(* IEC 61131-3 sources: sis-interlock-demo/tests/POUs/Generated/FB_VoteTruth_Test, 83 files *)

(* ---- FB_VoteTruth_Test.decl.st ---- *)
// AUTO-GENERATED by cemgen 1.0.0 — не редактировать: правьте матрицу и запустите
//   python -m cemgen generate <файл матрицы .csv или .xlsx>
// Матрица: SIS-V101-CEM, объект V-101, ревизия B от 2026-10-19, SHA-256 сетки df2ed4841a9453ca
// Назначение: набор coUnit: таблицы истинности голосования — F_VoteEval и FB_Voting по всем схемам,
//             политикам деградации и видам входа (DESIGN.md, 12.2). Экземпляр — GVL_TestsGenerated.
// Автор:      kr0nsch; код — генератор cemgen
// Версия:     1.0.0
// Документ:   docs/DESIGN.md, раздел «10. Генератор cemgen»; docs/cause_effect_matrix.md
// ВНИМАНИЕ:   код демонстрационный и не предназначен для систем безопасности. Реальная ПАЗ требует
//             определения SIL, сертифицированных аппаратных и программных средств и валидации по
//             ГОСТ Р МЭК 61511.
FUNCTION_BLOCK FB_VoteTruth_Test EXTENDS coUnit.FB_TestSuite
VAR
END_VAR

(* ---- ArchIndex.method.decl.st ---- *)
// AUTO-GENERATED by cemgen 1.0.0 — не редактировать: правьте матрицу и запустите
//   python -m cemgen generate <файл матрицы .csv или .xlsx>
// Матрица: SIS-V101-CEM, объект V-101, ревизия B от 2026-10-19, SHA-256 сетки df2ed4841a9453ca
// Назначение: вспомогательный метод набора FB_VoteTruth_Test.
// Автор:      kr0nsch; код — генератор cemgen
// Версия:     1.0.0
// Документ:   docs/DESIGN.md, раздел «10. Генератор cemgen»; docs/cause_effect_matrix.md
// ВНИМАНИЕ:   код демонстрационный и не предназначен для систем безопасности. Реальная ПАЗ требует
//             определения SIL, сертифицированных аппаратных и программных средств и валидации по
//             ГОСТ Р МЭК 61511.
// Индекс схемы в байте таблицы: 0 None, 1 1oo1, 2 1oo2, 3 2oo2, 4 2oo3, 5 ForcedTrip.
METHOD PRIVATE ArchIndex : BYTE
VAR_INPUT
    eArch : E_VoteArch;   // действующая схема
END_VAR

(* ---- ArchIndex.method.impl.st ---- *)
// AUTO-GENERATED by cemgen 1.0.0 — не редактировать: правьте матрицу и запустите
//   python -m cemgen generate <файл матрицы .csv или .xlsx>
// Матрица: SIS-V101-CEM, объект V-101, ревизия B от 2026-10-19, SHA-256 сетки df2ed4841a9453ca
CASE eArch OF
    E_VoteArch.Vote1oo1:
        ArchIndex := 1;
    E_VoteArch.Vote1oo2:
        ArchIndex := 2;
    E_VoteArch.Vote2oo2:
        ArchIndex := 3;
    E_VoteArch.Vote2oo3:
        ArchIndex := 4;
    E_VoteArch.ForcedTrip:
        ArchIndex := 5;
ELSE
    ArchIndex := 0;
END_CASE

(* ---- EncodeEval.method.decl.st ---- *)
// AUTO-GENERATED by cemgen 1.0.0 — не редактировать: правьте матрицу и запустите
//   python -m cemgen generate <файл матрицы .csv или .xlsx>
// Матрица: SIS-V101-CEM, объект V-101, ревизия B от 2026-10-19, SHA-256 сетки df2ed4841a9453ca
// Назначение: вспомогательный метод набора FB_VoteTruth_Test.
// Автор:      kr0nsch; код — генератор cemgen
// Версия:     1.0.0
// Документ:   docs/DESIGN.md, раздел «10. Генератор cemgen»; docs/cause_effect_matrix.md
// ВНИМАНИЕ:   код демонстрационный и не предназначен для систем безопасности. Реальная ПАЗ требует
//             определения SIL, сертифицированных аппаратных и программных средств и валидации по
//             ГОСТ Р МЭК 61511.
// Байт результата F_VoteEval: бит 0 — xTrip, бит 1 — xDegraded, биты 2–4 — индекс eArchEff.
METHOD PRIVATE EncodeEval : BYTE
VAR_INPUT
    stRes : ST_VoteResult;   // результат F_VoteEval
END_VAR

(* ---- EncodeFb.method.decl.st ---- *)
// AUTO-GENERATED by cemgen 1.0.0 — не редактировать: правьте матрицу и запустите
//   python -m cemgen generate <файл матрицы .csv или .xlsx>
// Матрица: SIS-V101-CEM, объект V-101, ревизия B от 2026-10-19, SHA-256 сетки df2ed4841a9453ca
// Назначение: вспомогательный метод набора FB_VoteTruth_Test.
// Автор:      kr0nsch; код — генератор cemgen
// Версия:     1.0.0
// Документ:   docs/DESIGN.md, раздел «10. Генератор cemgen»; docs/cause_effect_matrix.md
// ВНИМАНИЕ:   код демонстрационный и не предназначен для систем безопасности. Реальная ПАЗ требует
//             определения SIL, сертифицированных аппаратных и программных средств и валидации по
//             ГОСТ Р МЭК 61511.
// Байт результата FB_Voting: как у EncodeEval, плюс биты 5–7 — байпас каналов 1–3 в состоянии Active.
METHOD PRIVATE EncodeFb : BYTE
VAR_INPUT
    xTrip : BOOL;           // выход xTrip
    stSts : ST_VotingSts;   // состояние группы
END_VAR
VAR
    uiCh : UINT;            // канал
END_VAR

(* ---- EncodeFb.method.impl.st ---- *)
// AUTO-GENERATED by cemgen 1.0.0 — не редактировать: правьте матрицу и запустите
//   python -m cemgen generate <файл матрицы .csv или .xlsx>
// Матрица: SIS-V101-CEM, объект V-101, ревизия B от 2026-10-19, SHA-256 сетки df2ed4841a9453ca
EncodeFb := BOOL_TO_BYTE(xTrip) OR SHL(BOOL_TO_BYTE(stSts.xDegraded), 1)
    OR SHL(ArchIndex(eArch := stSts.eArchEff), 2);
FOR uiCh := 1 TO GVL_Const.SIS_VOTE_CH_MAX DO
    EncodeFb := EncodeFb OR SHL(BOOL_TO_BYTE(stSts.aeBypass[uiCh] = E_BypassState.Active), 4 + uiCh);
END_FOR

(* ---- Eval1oo1DAMatchesTable.method.decl.st ---- *)
// AUTO-GENERATED by cemgen 1.0.0 — не редактировать: правьте матрицу и запустите
//   python -m cemgen generate <файл матрицы .csv или .xlsx>
// Матрица: SIS-V101-CEM, объект V-101, ревизия B от 2026-10-19, SHA-256 сетки df2ed4841a9453ca
// Назначение: тест VoteTruth_Eval1oo1DA_MatchesTable набора FB_VoteTruth_Test.
// Автор:      kr0nsch; код — генератор cemgen
// Версия:     1.0.0
// Документ:   docs/DESIGN.md, раздел «10. Генератор cemgen»; docs/cause_effect_matrix.md
// ВНИМАНИЕ:   код демонстрационный и не предназначен для систем безопасности. Реальная ПАЗ требует
//             определения SIL, сертифицированных аппаратных и программных средств и валидации по
//             ГОСТ Р МЭК 61511.
// F_VoteEval, схема 1oo1, политика DegradeAvailable: все 4 сочетаний состояний каналов (Normal,
// Demand, Invalid, Bypassed) совпадают с таблицей TT_EVAL_1OO1_DA.
METHOD PRIVATE Eval1oo1DAMatchesTable
VAR
    uiRow      : UINT;                                                    // строка таблицы
    aeCh       : ARRAY[1..GVL_Const.SIS_VOTE_CH_MAX] OF E_ChannelState;   // состояния каналов строки
    stRes      : ST_VoteResult;                                           // результат F_VoteEval
    bAct       : BYTE;                                                    // фактический байт результата
    bExp       : BYTE;                                                    // ожидаемый байт из таблицы
    xMiss      : BOOL;                                                    // строка не совпала
    xFirst     : BOOL;                                                    // первая несовпавшая строка
    uiMismatch : UINT;                                                    // несовпавших строк
    uiFirstRow : UINT;                                                    // первая несовпавшая строка
    bFirstExp  : BYTE;                                                    // ожидаемый байт первой несовпавшей строки
    bFirstAct  : BYTE;                                                    // фактический байт первой несовпавшей строки
END_VAR

(* ---- Eval1oo1DAMatchesTable.method.impl.st ---- *)
// AUTO-GENERATED by cemgen 1.0.0 — не редактировать: правьте матрицу и запустите
//   python -m cemgen generate <файл матрицы .csv или .xlsx>
// Матрица: SIS-V101-CEM, объект V-101, ревизия B от 2026-10-19, SHA-256 сетки df2ed4841a9453ca
coUnit.TEST('VoteTruth_Eval1oo1DA_MatchesTable');
FOR uiRow := 0 TO 3 DO
    RowStates(uiRow := uiRow, uiChannels := 1, aeCh := aeCh);
    stRes := F_VoteEval(eArch := E_VoteArch.Vote1oo1, ePolicy := E_DegradePolicy.DegradeAvailable,
        aeCh := aeCh);
    bAct := EncodeEval(stRes := stRes);
    bExp := GVL_VoteTruthTable.TT_EVAL_1OO1_DA[uiRow];
    xMiss := bAct <> bExp;
    xFirst := xMiss AND uiMismatch = 0;
    uiFirstRow := SEL(xFirst, uiFirstRow, uiRow);
    bFirstExp := SEL(xFirst, bFirstExp, bExp);
    bFirstAct := SEL(xFirst, bFirstAct, bAct);
    uiMismatch := uiMismatch + BOOL_TO_UINT(xMiss);
END_FOR
AssertEquals_UINT(Expected := 0, Actual := uiMismatch,
    Message := MismatchText(sTable := 'TT_EVAL_1OO1_DA', uiRow := uiFirstRow, bExpected := bFirstExp,
        bActual := bFirstAct));
coUnit.TEST_FINISHED();

(* ---- Eval1oo1DSMatchesTable.method.decl.st ---- *)
// AUTO-GENERATED by cemgen 1.0.0 — не редактировать: правьте матрицу и запустите
//   python -m cemgen generate <файл матрицы .csv или .xlsx>
// Матрица: SIS-V101-CEM, объект V-101, ревизия B от 2026-10-19, SHA-256 сетки df2ed4841a9453ca
// Назначение: тест VoteTruth_Eval1oo1DS_MatchesTable набора FB_VoteTruth_Test.
// Автор:      kr0nsch; код — генератор cemgen
// Версия:     1.0.0
// Документ:   docs/DESIGN.md, раздел «10. Генератор cemgen»; docs/cause_effect_matrix.md
// ВНИМАНИЕ:   код демонстрационный и не предназначен для систем безопасности. Реальная ПАЗ требует
//             определения SIL, сертифицированных аппаратных и программных средств и валидации по
//             ГОСТ Р МЭК 61511.
// F_VoteEval, схема 1oo1, политика DegradeSafe: все 4 сочетаний состояний каналов (Normal, Demand,
// Invalid, Bypassed) совпадают с таблицей TT_EVAL_1OO1_DS.
METHOD PRIVATE Eval1oo1DSMatchesTable
VAR
    uiRow      : UINT;                                                    // строка таблицы
    aeCh       : ARRAY[1..GVL_Const.SIS_VOTE_CH_MAX] OF E_ChannelState;   // состояния каналов строки
    stRes      : ST_VoteResult;                                           // результат F_VoteEval
    bAct       : BYTE;                                                    // фактический байт результата
    bExp       : BYTE;                                                    // ожидаемый байт из таблицы
    xMiss      : BOOL;                                                    // строка не совпала
    xFirst     : BOOL;                                                    // первая несовпавшая строка
    uiMismatch : UINT;                                                    // несовпавших строк
    uiFirstRow : UINT;                                                    // первая несовпавшая строка
    bFirstExp  : BYTE;                                                    // ожидаемый байт первой несовпавшей строки
    bFirstAct  : BYTE;                                                    // фактический байт первой несовпавшей строки
END_VAR

(* ---- Eval1oo1DSMatchesTable.method.impl.st ---- *)
// AUTO-GENERATED by cemgen 1.0.0 — не редактировать: правьте матрицу и запустите
//   python -m cemgen generate <файл матрицы .csv или .xlsx>
// Матрица: SIS-V101-CEM, объект V-101, ревизия B от 2026-10-19, SHA-256 сетки df2ed4841a9453ca
coUnit.TEST('VoteTruth_Eval1oo1DS_MatchesTable');
FOR uiRow := 0 TO 3 DO
    RowStates(uiRow := uiRow, uiChannels := 1, aeCh := aeCh);
    stRes := F_VoteEval(eArch := E_VoteArch.Vote1oo1, ePolicy := E_DegradePolicy.DegradeSafe,
        aeCh := aeCh);
    bAct := EncodeEval(stRes := stRes);
    bExp := GVL_VoteTruthTable.TT_EVAL_1OO1_DS[uiRow];
    xMiss := bAct <> bExp;
    xFirst := xMiss AND uiMismatch = 0;
    uiFirstRow := SEL(xFirst, uiFirstRow, uiRow);
    bFirstExp := SEL(xFirst, bFirstExp, bExp);
    bFirstAct := SEL(xFirst, bFirstAct, bAct);
    uiMismatch := uiMismatch + BOOL_TO_UINT(xMiss);
END_FOR
AssertEquals_UINT(Expected := 0, Actual := uiMismatch,
    Message := MismatchText(sTable := 'TT_EVAL_1OO1_DS', uiRow := uiFirstRow, bExpected := bFirstExp,
        bActual := bFirstAct));
coUnit.TEST_FINISHED();

(* ---- Eval1oo1VTMatchesTable.method.decl.st ---- *)
// AUTO-GENERATED by cemgen 1.0.0 — не редактировать: правьте матрицу и запустите
//   python -m cemgen generate <файл матрицы .csv или .xlsx>
// Матрица: SIS-V101-CEM, объект V-101, ревизия B от 2026-10-19, SHA-256 сетки df2ed4841a9453ca
// Назначение: тест VoteTruth_Eval1oo1VT_MatchesTable набора FB_VoteTruth_Test.
// Автор:      kr0nsch; код — генератор cemgen
// Версия:     1.0.0
// Документ:   docs/DESIGN.md, раздел «10. Генератор cemgen»; docs/cause_effect_matrix.md
// ВНИМАНИЕ:   код демонстрационный и не предназначен для систем безопасности. Реальная ПАЗ требует
//             определения SIL, сертифицированных аппаратных и программных средств и валидации по
//             ГОСТ Р МЭК 61511.
// F_VoteEval, схема 1oo1, политика VoteTrip: все 4 сочетаний состояний каналов (Normal, Demand,
// Invalid, Bypassed) совпадают с таблицей TT_EVAL_1OO1_VT.
METHOD PRIVATE Eval1oo1VTMatchesTable
VAR
    uiRow      : UINT;                                                    // строка таблицы
    aeCh       : ARRAY[1..GVL_Const.SIS_VOTE_CH_MAX] OF E_ChannelState;   // состояния каналов строки
    stRes      : ST_VoteResult;                                           // результат F_VoteEval
    bAct       : BYTE;                                                    // фактический байт результата
    bExp       : BYTE;                                                    // ожидаемый байт из таблицы
    xMiss      : BOOL;                                                    // строка не совпала
    xFirst     : BOOL;                                                    // первая несовпавшая строка
    uiMismatch : UINT;                                                    // несовпавших строк
    uiFirstRow : UINT;                                                    // первая несовпавшая строка
    bFirstExp  : BYTE;                                                    // ожидаемый байт первой несовпавшей строки
    bFirstAct  : BYTE;                                                    // фактический байт первой несовпавшей строки
END_VAR

(* ---- Eval1oo1VTMatchesTable.method.impl.st ---- *)
// AUTO-GENERATED by cemgen 1.0.0 — не редактировать: правьте матрицу и запустите
//   python -m cemgen generate <файл матрицы .csv или .xlsx>
// Матрица: SIS-V101-CEM, объект V-101, ревизия B от 2026-10-19, SHA-256 сетки df2ed4841a9453ca
coUnit.TEST('VoteTruth_Eval1oo1VT_MatchesTable');
FOR uiRow := 0 TO 3 DO
    RowStates(uiRow := uiRow, uiChannels := 1, aeCh := aeCh);
    stRes := F_VoteEval(eArch := E_VoteArch.Vote1oo1, ePolicy := E_DegradePolicy.VoteTrip,
        aeCh := aeCh);
    bAct := EncodeEval(stRes := stRes);
    bExp := GVL_VoteTruthTable.TT_EVAL_1OO1_VT[uiRow];
    xMiss := bAct <> bExp;
    xFirst := xMiss AND uiMismatch = 0;
    uiFirstRow := SEL(xFirst, uiFirstRow, uiRow);
    bFirstExp := SEL(xFirst, bFirstExp, bExp);
    bFirstAct := SEL(xFirst, bFirstAct, bAct);
    uiMismatch := uiMismatch + BOOL_TO_UINT(xMiss);
END_FOR
AssertEquals_UINT(Expected := 0, Actual := uiMismatch,
    Message := MismatchText(sTable := 'TT_EVAL_1OO1_VT', uiRow := uiFirstRow, bExpected := bFirstExp,
        bActual := bFirstAct));
coUnit.TEST_FINISHED();

(* ---- Eval1oo2DAMatchesTable.method.decl.st ---- *)
// AUTO-GENERATED by cemgen 1.0.0 — не редактировать: правьте матрицу и запустите
//   python -m cemgen generate <файл матрицы .csv или .xlsx>
// Матрица: SIS-V101-CEM, объект V-101, ревизия B от 2026-10-19, SHA-256 сетки df2ed4841a9453ca
// Назначение: тест VoteTruth_Eval1oo2DA_MatchesTable набора FB_VoteTruth_Test.
// Автор:      kr0nsch; код — генератор cemgen
// Версия:     1.0.0
// Документ:   docs/DESIGN.md, раздел «10. Генератор cemgen»; docs/cause_effect_matrix.md
// ВНИМАНИЕ:   код демонстрационный и не предназначен для систем безопасности. Реальная ПАЗ требует
//             определения SIL, сертифицированных аппаратных и программных средств и валидации по
//             ГОСТ Р МЭК 61511.
// F_VoteEval, схема 1oo2, политика DegradeAvailable: все 16 сочетаний состояний каналов (Normal,
// Demand, Invalid, Bypassed) совпадают с таблицей TT_EVAL_1OO2_DA.
METHOD PRIVATE Eval1oo2DAMatchesTable
VAR
    uiRow      : UINT;                                                    // строка таблицы
    aeCh       : ARRAY[1..GVL_Const.SIS_VOTE_CH_MAX] OF E_ChannelState;   // состояния каналов строки
    stRes      : ST_VoteResult;                                           // результат F_VoteEval
    bAct       : BYTE;                                                    // фактический байт результата
    bExp       : BYTE;                                                    // ожидаемый байт из таблицы
    xMiss      : BOOL;                                                    // строка не совпала
    xFirst     : BOOL;                                                    // первая несовпавшая строка
    uiMismatch : UINT;                                                    // несовпавших строк
    uiFirstRow : UINT;                                                    // первая несовпавшая строка
    bFirstExp  : BYTE;                                                    // ожидаемый байт первой несовпавшей строки
    bFirstAct  : BYTE;                                                    // фактический байт первой несовпавшей строки
END_VAR

(* ---- Eval1oo2DAMatchesTable.method.impl.st ---- *)
// AUTO-GENERATED by cemgen 1.0.0 — не редактировать: правьте матрицу и запустите
//   python -m cemgen generate <файл матрицы .csv или .xlsx>
// Матрица: SIS-V101-CEM, объект V-101, ревизия B от 2026-10-19, SHA-256 сетки df2ed4841a9453ca
coUnit.TEST('VoteTruth_Eval1oo2DA_MatchesTable');
FOR uiRow := 0 TO 15 DO
    RowStates(uiRow := uiRow, uiChannels := 2, aeCh := aeCh);
    stRes := F_VoteEval(eArch := E_VoteArch.Vote1oo2, ePolicy := E_DegradePolicy.DegradeAvailable,
        aeCh := aeCh);
    bAct := EncodeEval(stRes := stRes);
    bExp := GVL_VoteTruthTable.TT_EVAL_1OO2_DA[uiRow];
    xMiss := bAct <> bExp;
    xFirst := xMiss AND uiMismatch = 0;
    uiFirstRow := SEL(xFirst, uiFirstRow, uiRow);
    bFirstExp := SEL(xFirst, bFirstExp, bExp);
    bFirstAct := SEL(xFirst, bFirstAct, bAct);
    uiMismatch := uiMismatch + BOOL_TO_UINT(xMiss);
END_FOR
AssertEquals_UINT(Expected := 0, Actual := uiMismatch,
    Message := MismatchText(sTable := 'TT_EVAL_1OO2_DA', uiRow := uiFirstRow, bExpected := bFirstExp,
        bActual := bFirstAct));
coUnit.TEST_FINISHED();

(* ---- Eval1oo2DSMatchesTable.method.decl.st ---- *)
// AUTO-GENERATED by cemgen 1.0.0 — не редактировать: правьте матрицу и запустите
//   python -m cemgen generate <файл матрицы .csv или .xlsx>
// Матрица: SIS-V101-CEM, объект V-101, ревизия B от 2026-10-19, SHA-256 сетки df2ed4841a9453ca
// Назначение: тест VoteTruth_Eval1oo2DS_MatchesTable набора FB_VoteTruth_Test.
// Автор:      kr0nsch; код — генератор cemgen
// Версия:     1.0.0
// Документ:   docs/DESIGN.md, раздел «10. Генератор cemgen»; docs/cause_effect_matrix.md
// ВНИМАНИЕ:   код демонстрационный и не предназначен для систем безопасности. Реальная ПАЗ требует
//             определения SIL, сертифицированных аппаратных и программных средств и валидации по
//             ГОСТ Р МЭК 61511.
// F_VoteEval, схема 1oo2, политика DegradeSafe: все 16 сочетаний состояний каналов (Normal, Demand,
// Invalid, Bypassed) совпадают с таблицей TT_EVAL_1OO2_DS.
METHOD PRIVATE Eval1oo2DSMatchesTable
VAR
    uiRow      : UINT;                                                    // строка таблицы
    aeCh       : ARRAY[1..GVL_Const.SIS_VOTE_CH_MAX] OF E_ChannelState;   // состояния каналов строки
    stRes      : ST_VoteResult;                                           // результат F_VoteEval
    bAct       : BYTE;                                                    // фактический байт результата
    bExp       : BYTE;                                                    // ожидаемый байт из таблицы
    xMiss      : BOOL;                                                    // строка не совпала
    xFirst     : BOOL;                                                    // первая несовпавшая строка
    uiMismatch : UINT;                                                    // несовпавших строк
    uiFirstRow : UINT;                                                    // первая несовпавшая строка
    bFirstExp  : BYTE;                                                    // ожидаемый байт первой несовпавшей строки
    bFirstAct  : BYTE;                                                    // фактический байт первой несовпавшей строки
END_VAR

(* ---- Eval1oo2DSMatchesTable.method.impl.st ---- *)
// AUTO-GENERATED by cemgen 1.0.0 — не редактировать: правьте матрицу и запустите
//   python -m cemgen generate <файл матрицы .csv или .xlsx>
// Матрица: SIS-V101-CEM, объект V-101, ревизия B от 2026-10-19, SHA-256 сетки df2ed4841a9453ca
coUnit.TEST('VoteTruth_Eval1oo2DS_MatchesTable');
FOR uiRow := 0 TO 15 DO
    RowStates(uiRow := uiRow, uiChannels := 2, aeCh := aeCh);
    stRes := F_VoteEval(eArch := E_VoteArch.Vote1oo2, ePolicy := E_DegradePolicy.DegradeSafe,
        aeCh := aeCh);
    bAct := EncodeEval(stRes := stRes);
    bExp := GVL_VoteTruthTable.TT_EVAL_1OO2_DS[uiRow];
    xMiss := bAct <> bExp;
    xFirst := xMiss AND uiMismatch = 0;
    uiFirstRow := SEL(xFirst, uiFirstRow, uiRow);
    bFirstExp := SEL(xFirst, bFirstExp, bExp);
    bFirstAct := SEL(xFirst, bFirstAct, bAct);
    uiMismatch := uiMismatch + BOOL_TO_UINT(xMiss);
END_FOR
AssertEquals_UINT(Expected := 0, Actual := uiMismatch,
    Message := MismatchText(sTable := 'TT_EVAL_1OO2_DS', uiRow := uiFirstRow, bExpected := bFirstExp,
        bActual := bFirstAct));
coUnit.TEST_FINISHED();

(* ---- Eval1oo2VTMatchesTable.method.decl.st ---- *)
// AUTO-GENERATED by cemgen 1.0.0 — не редактировать: правьте матрицу и запустите
//   python -m cemgen generate <файл матрицы .csv или .xlsx>
// Матрица: SIS-V101-CEM, объект V-101, ревизия B от 2026-10-19, SHA-256 сетки df2ed4841a9453ca
// Назначение: тест VoteTruth_Eval1oo2VT_MatchesTable набора FB_VoteTruth_Test.
// Автор:      kr0nsch; код — генератор cemgen
// Версия:     1.0.0
// Документ:   docs/DESIGN.md, раздел «10. Генератор cemgen»; docs/cause_effect_matrix.md
// ВНИМАНИЕ:   код демонстрационный и не предназначен для систем безопасности. Реальная ПАЗ требует
//             определения SIL, сертифицированных аппаратных и программных средств и валидации по
//             ГОСТ Р МЭК 61511.
// F_VoteEval, схема 1oo2, политика VoteTrip: все 16 сочетаний состояний каналов (Normal, Demand,
// Invalid, Bypassed) совпадают с таблицей TT_EVAL_1OO2_VT.
METHOD PRIVATE Eval1oo2VTMatchesTable
VAR
    uiRow      : UINT;                                                    // строка таблицы
    aeCh       : ARRAY[1..GVL_Const.SIS_VOTE_CH_MAX] OF E_ChannelState;   // состояния каналов строки
    stRes      : ST_VoteResult;                                           // результат F_VoteEval
    bAct       : BYTE;                                                    // фактический байт результата
    bExp       : BYTE;                                                    // ожидаемый байт из таблицы
    xMiss      : BOOL;                                                    // строка не совпала
    xFirst     : BOOL;                                                    // первая несовпавшая строка
    uiMismatch : UINT;                                                    // несовпавших строк
    uiFirstRow : UINT;                                                    // первая несовпавшая строка
    bFirstExp  : BYTE;                                                    // ожидаемый байт первой несовпавшей строки
    bFirstAct  : BYTE;                                                    // фактический байт первой несовпавшей строки
END_VAR

(* ---- Eval1oo2VTMatchesTable.method.impl.st ---- *)
// AUTO-GENERATED by cemgen 1.0.0 — не редактировать: правьте матрицу и запустите
//   python -m cemgen generate <файл матрицы .csv или .xlsx>
// Матрица: SIS-V101-CEM, объект V-101, ревизия B от 2026-10-19, SHA-256 сетки df2ed4841a9453ca
coUnit.TEST('VoteTruth_Eval1oo2VT_MatchesTable');
FOR uiRow := 0 TO 15 DO
    RowStates(uiRow := uiRow, uiChannels := 2, aeCh := aeCh);
    stRes := F_VoteEval(eArch := E_VoteArch.Vote1oo2, ePolicy := E_DegradePolicy.VoteTrip,
        aeCh := aeCh);
    bAct := EncodeEval(stRes := stRes);
    bExp := GVL_VoteTruthTable.TT_EVAL_1OO2_VT[uiRow];
    xMiss := bAct <> bExp;
    xFirst := xMiss AND uiMismatch = 0;
    uiFirstRow := SEL(xFirst, uiFirstRow, uiRow);
    bFirstExp := SEL(xFirst, bFirstExp, bExp);
    bFirstAct := SEL(xFirst, bFirstAct, bAct);
    uiMismatch := uiMismatch + BOOL_TO_UINT(xMiss);
END_FOR
AssertEquals_UINT(Expected := 0, Actual := uiMismatch,
    Message := MismatchText(sTable := 'TT_EVAL_1OO2_VT', uiRow := uiFirstRow, bExpected := bFirstExp,
        bActual := bFirstAct));
coUnit.TEST_FINISHED();

(* ---- Eval2oo2DAMatchesTable.method.decl.st ---- *)
// AUTO-GENERATED by cemgen 1.0.0 — не редактировать: правьте матрицу и запустите
//   python -m cemgen generate <файл матрицы .csv или .xlsx>
// Матрица: SIS-V101-CEM, объект V-101, ревизия B от 2026-10-19, SHA-256 сетки df2ed4841a9453ca
// Назначение: тест VoteTruth_Eval2oo2DA_MatchesTable набора FB_VoteTruth_Test.
// Автор:      kr0nsch; код — генератор cemgen
// Версия:     1.0.0
// Документ:   docs/DESIGN.md, раздел «10. Генератор cemgen»; docs/cause_effect_matrix.md
// ВНИМАНИЕ:   код демонстрационный и не предназначен для систем безопасности. Реальная ПАЗ требует
//             определения SIL, сертифицированных аппаратных и программных средств и валидации по
//             ГОСТ Р МЭК 61511.
// F_VoteEval, схема 2oo2, политика DegradeAvailable: все 16 сочетаний состояний каналов (Normal,
// Demand, Invalid, Bypassed) совпадают с таблицей TT_EVAL_2OO2_DA.
METHOD PRIVATE Eval2oo2DAMatchesTable
VAR
    uiRow      : UINT;                                                    // строка таблицы
    aeCh       : ARRAY[1..GVL_Const.SIS_VOTE_CH_MAX] OF E_ChannelState;   // состояния каналов строки
    stRes      : ST_VoteResult;                                           // результат F_VoteEval
    bAct       : BYTE;                                                    // фактический байт результата
    bExp       : BYTE;                                                    // ожидаемый байт из таблицы
    xMiss      : BOOL;                                                    // строка не совпала
    xFirst     : BOOL;                                                    // первая несовпавшая строка
    uiMismatch : UINT;                                                    // несовпавших строк
    uiFirstRow : UINT;                                                    // первая несовпавшая строка
    bFirstExp  : BYTE;                                                    // ожидаемый байт первой несовпавшей строки
    bFirstAct  : BYTE;                                                    // фактический байт первой несовпавшей строки
END_VAR

(* ---- Eval2oo2DAMatchesTable.method.impl.st ---- *)
// AUTO-GENERATED by cemgen 1.0.0 — не редактировать: правьте матрицу и запустите
//   python -m cemgen generate <файл матрицы .csv или .xlsx>
// Матрица: SIS-V101-CEM, объект V-101, ревизия B от 2026-10-19, SHA-256 сетки df2ed4841a9453ca
coUnit.TEST('VoteTruth_Eval2oo2DA_MatchesTable');
FOR uiRow := 0 TO 15 DO
    RowStates(uiRow := uiRow, uiChannels := 2, aeCh := aeCh);
    stRes := F_VoteEval(eArch := E_VoteArch.Vote2oo2, ePolicy := E_DegradePolicy.DegradeAvailable,
        aeCh := aeCh);
    bAct := EncodeEval(stRes := stRes);
    bExp := GVL_VoteTruthTable.TT_EVAL_2OO2_DA[uiRow];
    xMiss := bAct <> bExp;
    xFirst := xMiss AND uiMismatch = 0;
    uiFirstRow := SEL(xFirst, uiFirstRow, uiRow);
    bFirstExp := SEL(xFirst, bFirstExp, bExp);
    bFirstAct := SEL(xFirst, bFirstAct, bAct);
    uiMismatch := uiMismatch + BOOL_TO_UINT(xMiss);
END_FOR
AssertEquals_UINT(Expected := 0, Actual := uiMismatch,
    Message := MismatchText(sTable := 'TT_EVAL_2OO2_DA', uiRow := uiFirstRow, bExpected := bFirstExp,
        bActual := bFirstAct));
coUnit.TEST_FINISHED();

(* ---- Eval2oo2DSMatchesTable.method.decl.st ---- *)
// AUTO-GENERATED by cemgen 1.0.0 — не редактировать: правьте матрицу и запустите
//   python -m cemgen generate <файл матрицы .csv или .xlsx>
// Матрица: SIS-V101-CEM, объект V-101, ревизия B от 2026-10-19, SHA-256 сетки df2ed4841a9453ca
// Назначение: тест VoteTruth_Eval2oo2DS_MatchesTable набора FB_VoteTruth_Test.
// Автор:      kr0nsch; код — генератор cemgen
// Версия:     1.0.0
// Документ:   docs/DESIGN.md, раздел «10. Генератор cemgen»; docs/cause_effect_matrix.md
// ВНИМАНИЕ:   код демонстрационный и не предназначен для систем безопасности. Реальная ПАЗ требует
//             определения SIL, сертифицированных аппаратных и программных средств и валидации по
//             ГОСТ Р МЭК 61511.
// F_VoteEval, схема 2oo2, политика DegradeSafe: все 16 сочетаний состояний каналов (Normal, Demand,
// Invalid, Bypassed) совпадают с таблицей TT_EVAL_2OO2_DS.
METHOD PRIVATE Eval2oo2DSMatchesTable
VAR
    uiRow      : UINT;                                                    // строка таблицы
    aeCh       : ARRAY[1..GVL_Const.SIS_VOTE_CH_MAX] OF E_ChannelState;   // состояния каналов строки
    stRes      : ST_VoteResult;                                           // результат F_VoteEval
    bAct       : BYTE;                                                    // фактический байт результата
    bExp       : BYTE;                                                    // ожидаемый байт из таблицы
    xMiss      : BOOL;                                                    // строка не совпала
    xFirst     : BOOL;                                                    // первая несовпавшая строка
    uiMismatch : UINT;                                                    // несовпавших строк
    uiFirstRow : UINT;                                                    // первая несовпавшая строка
    bFirstExp  : BYTE;                                                    // ожидаемый байт первой несовпавшей строки
    bFirstAct  : BYTE;                                                    // фактический байт первой несовпавшей строки
END_VAR

(* ---- Eval2oo2DSMatchesTable.method.impl.st ---- *)
// AUTO-GENERATED by cemgen 1.0.0 — не редактировать: правьте матрицу и запустите
//   python -m cemgen generate <файл матрицы .csv или .xlsx>
// Матрица: SIS-V101-CEM, объект V-101, ревизия B от 2026-10-19, SHA-256 сетки df2ed4841a9453ca
coUnit.TEST('VoteTruth_Eval2oo2DS_MatchesTable');
FOR uiRow := 0 TO 15 DO
    RowStates(uiRow := uiRow, uiChannels := 2, aeCh := aeCh);
    stRes := F_VoteEval(eArch := E_VoteArch.Vote2oo2, ePolicy := E_DegradePolicy.DegradeSafe,
        aeCh := aeCh);
    bAct := EncodeEval(stRes := stRes);
    bExp := GVL_VoteTruthTable.TT_EVAL_2OO2_DS[uiRow];
    xMiss := bAct <> bExp;
    xFirst := xMiss AND uiMismatch = 0;
    uiFirstRow := SEL(xFirst, uiFirstRow, uiRow);
    bFirstExp := SEL(xFirst, bFirstExp, bExp);
    bFirstAct := SEL(xFirst, bFirstAct, bAct);
    uiMismatch := uiMismatch + BOOL_TO_UINT(xMiss);
END_FOR
AssertEquals_UINT(Expected := 0, Actual := uiMismatch,
    Message := MismatchText(sTable := 'TT_EVAL_2OO2_DS', uiRow := uiFirstRow, bExpected := bFirstExp,
        bActual := bFirstAct));
coUnit.TEST_FINISHED();

(* ---- Eval2oo2VTMatchesTable.method.decl.st ---- *)
// AUTO-GENERATED by cemgen 1.0.0 — не редактировать: правьте матрицу и запустите
//   python -m cemgen generate <файл матрицы .csv или .xlsx>
// Матрица: SIS-V101-CEM, объект V-101, ревизия B от 2026-10-19, SHA-256 сетки df2ed4841a9453ca
// Назначение: тест VoteTruth_Eval2oo2VT_MatchesTable набора FB_VoteTruth_Test.
// Автор:      kr0nsch; код — генератор cemgen
// Версия:     1.0.0
// Документ:   docs/DESIGN.md, раздел «10. Генератор cemgen»; docs/cause_effect_matrix.md
// ВНИМАНИЕ:   код демонстрационный и не предназначен для систем безопасности. Реальная ПАЗ требует
//             определения SIL, сертифицированных аппаратных и программных средств и валидации по
//             ГОСТ Р МЭК 61511.
// F_VoteEval, схема 2oo2, политика VoteTrip: все 16 сочетаний состояний каналов (Normal, Demand,
// Invalid, Bypassed) совпадают с таблицей TT_EVAL_2OO2_VT.
METHOD PRIVATE Eval2oo2VTMatchesTable
VAR
    uiRow      : UINT;                                                    // строка таблицы
    aeCh       : ARRAY[1..GVL_Const.SIS_VOTE_CH_MAX] OF E_ChannelState;   // состояния каналов строки
    stRes      : ST_VoteResult;                                           // результат F_VoteEval
    bAct       : BYTE;                                                    // фактический байт результата
    bExp       : BYTE;                                                    // ожидаемый байт из таблицы
    xMiss      : BOOL;                                                    // строка не совпала
    xFirst     : BOOL;                                                    // первая несовпавшая строка
    uiMismatch : UINT;                                                    // несовпавших строк
    uiFirstRow : UINT;                                                    // первая несовпавшая строка
    bFirstExp  : BYTE;                                                    // ожидаемый байт первой несовпавшей строки
    bFirstAct  : BYTE;                                                    // фактический байт первой несовпавшей строки
END_VAR

(* ---- Eval2oo2VTMatchesTable.method.impl.st ---- *)
// AUTO-GENERATED by cemgen 1.0.0 — не редактировать: правьте матрицу и запустите
//   python -m cemgen generate <файл матрицы .csv или .xlsx>
// Матрица: SIS-V101-CEM, объект V-101, ревизия B от 2026-10-19, SHA-256 сетки df2ed4841a9453ca
coUnit.TEST('VoteTruth_Eval2oo2VT_MatchesTable');
FOR uiRow := 0 TO 15 DO
    RowStates(uiRow := uiRow, uiChannels := 2, aeCh := aeCh);
    stRes := F_VoteEval(eArch := E_VoteArch.Vote2oo2, ePolicy := E_DegradePolicy.VoteTrip,
        aeCh := aeCh);
    bAct := EncodeEval(stRes := stRes);
    bExp := GVL_VoteTruthTable.TT_EVAL_2OO2_VT[uiRow];
    xMiss := bAct <> bExp;
    xFirst := xMiss AND uiMismatch = 0;
    uiFirstRow := SEL(xFirst, uiFirstRow, uiRow);
    bFirstExp := SEL(xFirst, bFirstExp, bExp);
    bFirstAct := SEL(xFirst, bFirstAct, bAct);
    uiMismatch := uiMismatch + BOOL_TO_UINT(xMiss);
END_FOR
AssertEquals_UINT(Expected := 0, Actual := uiMismatch,
    Message := MismatchText(sTable := 'TT_EVAL_2OO2_VT', uiRow := uiFirstRow, bExpected := bFirstExp,
        bActual := bFirstAct));
coUnit.TEST_FINISHED();

(* ---- Eval2oo3DAMatchesTable.method.decl.st ---- *)
// AUTO-GENERATED by cemgen 1.0.0 — не редактировать: правьте матрицу и запустите
//   python -m cemgen generate <файл матрицы .csv или .xlsx>
// Матрица: SIS-V101-CEM, объект V-101, ревизия B от 2026-10-19, SHA-256 сетки df2ed4841a9453ca
// Назначение: тест VoteTruth_Eval2oo3DA_MatchesTable набора FB_VoteTruth_Test.
// Автор:      kr0nsch; код — генератор cemgen
// Версия:     1.0.0
// Документ:   docs/DESIGN.md, раздел «10. Генератор cemgen»; docs/cause_effect_matrix.md
// ВНИМАНИЕ:   код демонстрационный и не предназначен для систем безопасности. Реальная ПАЗ требует
//             определения SIL, сертифицированных аппаратных и программных средств и валидации по
//             ГОСТ Р МЭК 61511.
// F_VoteEval, схема 2oo3, политика DegradeAvailable: все 64 сочетаний состояний каналов (Normal,
// Demand, Invalid, Bypassed) совпадают с таблицей TT_EVAL_2OO3_DA.
METHOD PRIVATE Eval2oo3DAMatchesTable
VAR
    uiRow      : UINT;                                                    // строка таблицы
    aeCh       : ARRAY[1..GVL_Const.SIS_VOTE_CH_MAX] OF E_ChannelState;   // состояния каналов строки
    stRes      : ST_VoteResult;                                           // результат F_VoteEval
    bAct       : BYTE;                                                    // фактический байт результата
    bExp       : BYTE;                                                    // ожидаемый байт из таблицы
    xMiss      : BOOL;                                                    // строка не совпала
    xFirst     : BOOL;                                                    // первая несовпавшая строка
    uiMismatch : UINT;                                                    // несовпавших строк
    uiFirstRow : UINT;                                                    // первая несовпавшая строка
    bFirstExp  : BYTE;                                                    // ожидаемый байт первой несовпавшей строки
    bFirstAct  : BYTE;                                                    // фактический байт первой несовпавшей строки
END_VAR

(* ---- Eval2oo3DAMatchesTable.method.impl.st ---- *)
// AUTO-GENERATED by cemgen 1.0.0 — не редактировать: правьте матрицу и запустите
//   python -m cemgen generate <файл матрицы .csv или .xlsx>
// Матрица: SIS-V101-CEM, объект V-101, ревизия B от 2026-10-19, SHA-256 сетки df2ed4841a9453ca
coUnit.TEST('VoteTruth_Eval2oo3DA_MatchesTable');
FOR uiRow := 0 TO 63 DO
    RowStates(uiRow := uiRow, uiChannels := 3, aeCh := aeCh);
    stRes := F_VoteEval(eArch := E_VoteArch.Vote2oo3, ePolicy := E_DegradePolicy.DegradeAvailable,
        aeCh := aeCh);
    bAct := EncodeEval(stRes := stRes);
    bExp := GVL_VoteTruthTable.TT_EVAL_2OO3_DA[uiRow];
    xMiss := bAct <> bExp;
    xFirst := xMiss AND uiMismatch = 0;
    uiFirstRow := SEL(xFirst, uiFirstRow, uiRow);
    bFirstExp := SEL(xFirst, bFirstExp, bExp);
    bFirstAct := SEL(xFirst, bFirstAct, bAct);
    uiMismatch := uiMismatch + BOOL_TO_UINT(xMiss);
END_FOR
AssertEquals_UINT(Expected := 0, Actual := uiMismatch,
    Message := MismatchText(sTable := 'TT_EVAL_2OO3_DA', uiRow := uiFirstRow, bExpected := bFirstExp,
        bActual := bFirstAct));
coUnit.TEST_FINISHED();

(* ---- Eval2oo3DSMatchesTable.method.decl.st ---- *)
// AUTO-GENERATED by cemgen 1.0.0 — не редактировать: правьте матрицу и запустите
//   python -m cemgen generate <файл матрицы .csv или .xlsx>
// Матрица: SIS-V101-CEM, объект V-101, ревизия B от 2026-10-19, SHA-256 сетки df2ed4841a9453ca
// Назначение: тест VoteTruth_Eval2oo3DS_MatchesTable набора FB_VoteTruth_Test.
// Автор:      kr0nsch; код — генератор cemgen
// Версия:     1.0.0
// Документ:   docs/DESIGN.md, раздел «10. Генератор cemgen»; docs/cause_effect_matrix.md
// ВНИМАНИЕ:   код демонстрационный и не предназначен для систем безопасности. Реальная ПАЗ требует
//             определения SIL, сертифицированных аппаратных и программных средств и валидации по
//             ГОСТ Р МЭК 61511.
// F_VoteEval, схема 2oo3, политика DegradeSafe: все 64 сочетаний состояний каналов (Normal, Demand,
// Invalid, Bypassed) совпадают с таблицей TT_EVAL_2OO3_DS.
METHOD PRIVATE Eval2oo3DSMatchesTable
VAR
    uiRow      : UINT;                                                    // строка таблицы
    aeCh       : ARRAY[1..GVL_Const.SIS_VOTE_CH_MAX] OF E_ChannelState;   // состояния каналов строки
    stRes      : ST_VoteResult;                                           // результат F_VoteEval
    bAct       : BYTE;                                                    // фактический байт результата
    bExp       : BYTE;                                                    // ожидаемый байт из таблицы
    xMiss      : BOOL;                                                    // строка не совпала
    xFirst     : BOOL;                                                    // первая несовпавшая строка
    uiMismatch : UINT;                                                    // несовпавших строк
    uiFirstRow : UINT;                                                    // первая несовпавшая строка
    bFirstExp  : BYTE;                                                    // ожидаемый байт первой несовпавшей строки
    bFirstAct  : BYTE;                                                    // фактический байт первой несовпавшей строки
END_VAR

(* ---- Eval2oo3DSMatchesTable.method.impl.st ---- *)
// AUTO-GENERATED by cemgen 1.0.0 — не редактировать: правьте матрицу и запустите
//   python -m cemgen generate <файл матрицы .csv или .xlsx>
// Матрица: SIS-V101-CEM, объект V-101, ревизия B от 2026-10-19, SHA-256 сетки df2ed4841a9453ca
coUnit.TEST('VoteTruth_Eval2oo3DS_MatchesTable');
FOR uiRow := 0 TO 63 DO
    RowStates(uiRow := uiRow, uiChannels := 3, aeCh := aeCh);
    stRes := F_VoteEval(eArch := E_VoteArch.Vote2oo3, ePolicy := E_DegradePolicy.DegradeSafe,
        aeCh := aeCh);
    bAct := EncodeEval(stRes := stRes);
    bExp := GVL_VoteTruthTable.TT_EVAL_2OO3_DS[uiRow];
    xMiss := bAct <> bExp;
    xFirst := xMiss AND uiMismatch = 0;
    uiFirstRow := SEL(xFirst, uiFirstRow, uiRow);
    bFirstExp := SEL(xFirst, bFirstExp, bExp);
    bFirstAct := SEL(xFirst, bFirstAct, bAct);
    uiMismatch := uiMismatch + BOOL_TO_UINT(xMiss);
END_FOR
AssertEquals_UINT(Expected := 0, Actual := uiMismatch,
    Message := MismatchText(sTable := 'TT_EVAL_2OO3_DS', uiRow := uiFirstRow, bExpected := bFirstExp,
        bActual := bFirstAct));
coUnit.TEST_FINISHED();

(* ---- Eval2oo3VTMatchesTable.method.decl.st ---- *)
// AUTO-GENERATED by cemgen 1.0.0 — не редактировать: правьте матрицу и запустите
//   python -m cemgen generate <файл матрицы .csv или .xlsx>
// Матрица: SIS-V101-CEM, объект V-101, ревизия B от 2026-10-19, SHA-256 сетки df2ed4841a9453ca
// Назначение: тест VoteTruth_Eval2oo3VT_MatchesTable набора FB_VoteTruth_Test.
// Автор:      kr0nsch; код — генератор cemgen
// Версия:     1.0.0
// Документ:   docs/DESIGN.md, раздел «10. Генератор cemgen»; docs/cause_effect_matrix.md
// ВНИМАНИЕ:   код демонстрационный и не предназначен для систем безопасности. Реальная ПАЗ требует
//             определения SIL, сертифицированных аппаратных и программных средств и валидации по
//             ГОСТ Р МЭК 61511.
// F_VoteEval, схема 2oo3, политика VoteTrip: все 64 сочетаний состояний каналов (Normal, Demand,
// Invalid, Bypassed) совпадают с таблицей TT_EVAL_2OO3_VT.
METHOD PRIVATE Eval2oo3VTMatchesTable
VAR
    uiRow      : UINT;                                                    // строка таблицы
    aeCh       : ARRAY[1..GVL_Const.SIS_VOTE_CH_MAX] OF E_ChannelState;   // состояния каналов строки
    stRes      : ST_VoteResult;                                           // результат F_VoteEval
    bAct       : BYTE;                                                    // фактический байт результата
    bExp       : BYTE;                                                    // ожидаемый байт из таблицы
    xMiss      : BOOL;                                                    // строка не совпала
    xFirst     : BOOL;                                                    // первая несовпавшая строка
    uiMismatch : UINT;                                                    // несовпавших строк
    uiFirstRow : UINT;                                                    // первая несовпавшая строка
    bFirstExp  : BYTE;                                                    // ожидаемый байт первой несовпавшей строки
    bFirstAct  : BYTE;                                                    // фактический байт первой несовпавшей строки
END_VAR

(* ---- Eval2oo3VTMatchesTable.method.impl.st ---- *)
// AUTO-GENERATED by cemgen 1.0.0 — не редактировать: правьте матрицу и запустите
//   python -m cemgen generate <файл матрицы .csv или .xlsx>
// Матрица: SIS-V101-CEM, объект V-101, ревизия B от 2026-10-19, SHA-256 сетки df2ed4841a9453ca
coUnit.TEST('VoteTruth_Eval2oo3VT_MatchesTable');
FOR uiRow := 0 TO 63 DO
    RowStates(uiRow := uiRow, uiChannels := 3, aeCh := aeCh);
    stRes := F_VoteEval(eArch := E_VoteArch.Vote2oo3, ePolicy := E_DegradePolicy.VoteTrip,
        aeCh := aeCh);
    bAct := EncodeEval(stRes := stRes);
    bExp := GVL_VoteTruthTable.TT_EVAL_2OO3_VT[uiRow];
    xMiss := bAct <> bExp;
    xFirst := xMiss AND uiMismatch = 0;
    uiFirstRow := SEL(xFirst, uiFirstRow, uiRow);
    bFirstExp := SEL(xFirst, bFirstExp, bExp);
    bFirstAct := SEL(xFirst, bFirstAct, bAct);
    uiMismatch := uiMismatch + BOOL_TO_UINT(xMiss);
END_FOR
AssertEquals_UINT(Expected := 0, Actual := uiMismatch,
    Message := MismatchText(sTable := 'TT_EVAL_2OO3_VT', uiRow := uiFirstRow, bExpected := bFirstExp,
        bActual := bFirstAct));
coUnit.TEST_FINISHED();

(* ---- Fb1oo1DAAIMatchesTable.method.decl.st ---- *)
// AUTO-GENERATED by cemgen 1.0.0 — не редактировать: правьте матрицу и запустите
//   python -m cemgen generate <файл матрицы .csv или .xlsx>
// Матрица: SIS-V101-CEM, объект V-101, ревизия B от 2026-10-19, SHA-256 сетки df2ed4841a9453ca
// Назначение: тест VoteTruth_Fb1oo1DAAI_MatchesTable набора FB_VoteTruth_Test.
// Автор:      kr0nsch; код — генератор cemgen
// Версия:     1.0.0
// Документ:   docs/DESIGN.md, раздел «10. Генератор cemgen»; docs/cause_effect_matrix.md
// ВНИМАНИЕ:   код демонстрационный и не предназначен для систем безопасности. Реальная ПАЗ требует
//             определения SIL, сертифицированных аппаратных и программных средств и валидации по
//             ГОСТ Р МЭК 61511.
// FB_Voting, схема 1oo1, политика DegradeAvailable, аналоговые каналы: все 8 сочетаний «требование ×
// достоверность × запрос байпаса» совпадают с таблицей TT_FB_1OO1_DA_AI. На строку — два вызова одного
// экземпляра: без запросов байпаса (сброс байпасов прошлой строки) и с полной строкой.
METHOD PRIVATE Fb1oo1DAAIMatchesTable
VAR
    fbTime     : PL.FB_FakeTime;   // время не меняется
    fbVote     : FB_Voting;        // ФБ под тестом, один экземпляр на все строки
    stCfg      : ST_VotingCfg;     // конфигурация теста уровня 2
    stIn       : ST_VoteIn;        // входы строки
    stCmd      : ST_VoteCmd;       // запросы байпаса строки
    uiRow      : UINT;             // строка таблицы
    bAct       : BYTE;             // фактический байт результата
    bExp       : BYTE;             // ожидаемый байт из таблицы
    xMiss      : BOOL;             // строка не совпала
    xFirst     : BOOL;             // первая несовпавшая строка
    uiMismatch : UINT;             // несовпавших строк
    uiFirstRow : UINT;             // первая несовпавшая строка
    bFirstExp  : BYTE;             // ожидаемый байт первой несовпавшей строки
    bFirstAct  : BYTE;             // фактический байт первой несовпавшей строки
END_VAR

(* ---- Fb1oo1DAAIMatchesTable.method.impl.st ---- *)
// AUTO-GENERATED by cemgen 1.0.0 — не редактировать: правьте матрицу и запустите
//   python -m cemgen generate <файл матрицы .csv или .xlsx>
// Матрица: SIS-V101-CEM, объект V-101, ревизия B от 2026-10-19, SHA-256 сетки df2ed4841a9453ca
coUnit.TEST('VoteTruth_Fb1oo1DAAI_MatchesTable');
stCfg.eArch := E_VoteArch.Vote1oo1;
stCfg.ePolicy := E_DegradePolicy.DegradeAvailable;
stCfg.eInput := E_SisInputKind.Analog;
stCfg.xDiHealthy := TRUE;
stCfg.eLimitDir := E_LimitDir.High;
stCfg.rTripLimit_eu := 50.0;
stCfg.rHyst_eu := 0.0;
stCfg.rDiscrepancyMax_eu := 0.0;
stCfg.tDiscrepancyDelay := T#0S;
stCfg.tBypassMax := T#1H;
stCfg.uiMaxBypass := 0;
FOR uiRow := 0 TO 7 DO
    RowInputs(uiRow := uiRow, uiChannels := 1, xBypass := FALSE, stIn := stIn, stCmd := stCmd);
    fbVote(stIn := stIn, stCmd := stCmd, stCfg := stCfg, xBypassPermit := TRUE, uiCause := 1,
        itfTime := fbTime);
    RowInputs(uiRow := uiRow, uiChannels := 1, xBypass := TRUE, stIn := stIn, stCmd := stCmd);
    fbVote(stIn := stIn, stCmd := stCmd, stCfg := stCfg, xBypassPermit := TRUE, uiCause := 1,
        itfTime := fbTime);
    bAct := EncodeFb(xTrip := fbVote.xTrip, stSts := fbVote.stSts);
    bExp := GVL_VoteTruthTable.TT_FB_1OO1_DA_AI[uiRow];
    xMiss := bAct <> bExp;
    xFirst := xMiss AND uiMismatch = 0;
    uiFirstRow := SEL(xFirst, uiFirstRow, uiRow);
    bFirstExp := SEL(xFirst, bFirstExp, bExp);
    bFirstAct := SEL(xFirst, bFirstAct, bAct);
    uiMismatch := uiMismatch + BOOL_TO_UINT(xMiss);
END_FOR
AssertEquals_UINT(Expected := 0, Actual := uiMismatch,
    Message := MismatchText(sTable := 'TT_FB_1OO1_DA_AI', uiRow := uiFirstRow, bExpected := bFirstExp,
        bActual := bFirstAct));
coUnit.TEST_FINISHED();

(* ---- Fb1oo1DADIMatchesTable.method.decl.st ---- *)
// AUTO-GENERATED by cemgen 1.0.0 — не редактировать: правьте матрицу и запустите
//   python -m cemgen generate <файл матрицы .csv или .xlsx>
// Матрица: SIS-V101-CEM, объект V-101, ревизия B от 2026-10-19, SHA-256 сетки df2ed4841a9453ca
// Назначение: тест VoteTruth_Fb1oo1DADI_MatchesTable набора FB_VoteTruth_Test.
// Автор:      kr0nsch; код — генератор cemgen
// Версия:     1.0.0
// Документ:   docs/DESIGN.md, раздел «10. Генератор cemgen»; docs/cause_effect_matrix.md
// ВНИМАНИЕ:   код демонстрационный и не предназначен для систем безопасности. Реальная ПАЗ требует
//             определения SIL, сертифицированных аппаратных и программных средств и валидации по
//             ГОСТ Р МЭК 61511.
// FB_Voting, схема 1oo1, политика DegradeAvailable, дискретные каналы: все 8 сочетаний «требование ×
// достоверность × запрос байпаса» совпадают с таблицей TT_FB_1OO1_DA_DI. На строку — два вызова одного
// экземпляра: без запросов байпаса (сброс байпасов прошлой строки) и с полной строкой.
METHOD PRIVATE Fb1oo1DADIMatchesTable
VAR
    fbTime     : PL.FB_FakeTime;   // время не меняется
    fbVote     : FB_Voting;        // ФБ под тестом, один экземпляр на все строки
    stCfg      : ST_VotingCfg;     // конфигурация теста уровня 2
    stIn       : ST_VoteIn;        // входы строки
    stCmd      : ST_VoteCmd;       // запросы байпаса строки
    uiRow      : UINT;             // строка таблицы
    bAct       : BYTE;             // фактический байт результата
    bExp       : BYTE;             // ожидаемый байт из таблицы
    xMiss      : BOOL;             // строка не совпала
    xFirst     : BOOL;             // первая несовпавшая строка
    uiMismatch : UINT;             // несовпавших строк
    uiFirstRow : UINT;             // первая несовпавшая строка
    bFirstExp  : BYTE;             // ожидаемый байт первой несовпавшей строки
    bFirstAct  : BYTE;             // фактический байт первой несовпавшей строки
END_VAR

(* ---- Fb1oo1DADIMatchesTable.method.impl.st ---- *)
// AUTO-GENERATED by cemgen 1.0.0 — не редактировать: правьте матрицу и запустите
//   python -m cemgen generate <файл матрицы .csv или .xlsx>
// Матрица: SIS-V101-CEM, объект V-101, ревизия B от 2026-10-19, SHA-256 сетки df2ed4841a9453ca
coUnit.TEST('VoteTruth_Fb1oo1DADI_MatchesTable');
stCfg.eArch := E_VoteArch.Vote1oo1;
stCfg.ePolicy := E_DegradePolicy.DegradeAvailable;
stCfg.eInput := E_SisInputKind.Discrete;
stCfg.xDiHealthy := TRUE;
stCfg.eLimitDir := E_LimitDir.High;
stCfg.rTripLimit_eu := 50.0;
stCfg.rHyst_eu := 0.0;
stCfg.rDiscrepancyMax_eu := 0.0;
stCfg.tDiscrepancyDelay := T#0S;
stCfg.tBypassMax := T#1H;
stCfg.uiMaxBypass := 0;
FOR uiRow := 0 TO 7 DO
    RowInputs(uiRow := uiRow, uiChannels := 1, xBypass := FALSE, stIn := stIn, stCmd := stCmd);
    fbVote(stIn := stIn, stCmd := stCmd, stCfg := stCfg, xBypassPermit := TRUE, uiCause := 1,
        itfTime := fbTime);
    RowInputs(uiRow := uiRow, uiChannels := 1, xBypass := TRUE, stIn := stIn, stCmd := stCmd);
    fbVote(stIn := stIn, stCmd := stCmd, stCfg := stCfg, xBypassPermit := TRUE, uiCause := 1,
        itfTime := fbTime);
    bAct := EncodeFb(xTrip := fbVote.xTrip, stSts := fbVote.stSts);
    bExp := GVL_VoteTruthTable.TT_FB_1OO1_DA_DI[uiRow];
    xMiss := bAct <> bExp;
    xFirst := xMiss AND uiMismatch = 0;
    uiFirstRow := SEL(xFirst, uiFirstRow, uiRow);
    bFirstExp := SEL(xFirst, bFirstExp, bExp);
    bFirstAct := SEL(xFirst, bFirstAct, bAct);
    uiMismatch := uiMismatch + BOOL_TO_UINT(xMiss);
END_FOR
AssertEquals_UINT(Expected := 0, Actual := uiMismatch,
    Message := MismatchText(sTable := 'TT_FB_1OO1_DA_DI', uiRow := uiFirstRow, bExpected := bFirstExp,
        bActual := bFirstAct));
coUnit.TEST_FINISHED();

(* ---- Fb1oo1DSAIMatchesTable.method.decl.st ---- *)
// AUTO-GENERATED by cemgen 1.0.0 — не редактировать: правьте матрицу и запустите
//   python -m cemgen generate <файл матрицы .csv или .xlsx>
// Матрица: SIS-V101-CEM, объект V-101, ревизия B от 2026-10-19, SHA-256 сетки df2ed4841a9453ca
// Назначение: тест VoteTruth_Fb1oo1DSAI_MatchesTable набора FB_VoteTruth_Test.
// Автор:      kr0nsch; код — генератор cemgen
// Версия:     1.0.0
// Документ:   docs/DESIGN.md, раздел «10. Генератор cemgen»; docs/cause_effect_matrix.md
// ВНИМАНИЕ:   код демонстрационный и не предназначен для систем безопасности. Реальная ПАЗ требует
//             определения SIL, сертифицированных аппаратных и программных средств и валидации по
//             ГОСТ Р МЭК 61511.
// FB_Voting, схема 1oo1, политика DegradeSafe, аналоговые каналы: все 8 сочетаний «требование ×
// достоверность × запрос байпаса» совпадают с таблицей TT_FB_1OO1_DS_AI. На строку — два вызова одного
// экземпляра: без запросов байпаса (сброс байпасов прошлой строки) и с полной строкой.
METHOD PRIVATE Fb1oo1DSAIMatchesTable
VAR
    fbTime     : PL.FB_FakeTime;   // время не меняется
    fbVote     : FB_Voting;        // ФБ под тестом, один экземпляр на все строки
    stCfg      : ST_VotingCfg;     // конфигурация теста уровня 2
    stIn       : ST_VoteIn;        // входы строки
    stCmd      : ST_VoteCmd;       // запросы байпаса строки
    uiRow      : UINT;             // строка таблицы
    bAct       : BYTE;             // фактический байт результата
    bExp       : BYTE;             // ожидаемый байт из таблицы
    xMiss      : BOOL;             // строка не совпала
    xFirst     : BOOL;             // первая несовпавшая строка
    uiMismatch : UINT;             // несовпавших строк
    uiFirstRow : UINT;             // первая несовпавшая строка
    bFirstExp  : BYTE;             // ожидаемый байт первой несовпавшей строки
    bFirstAct  : BYTE;             // фактический байт первой несовпавшей строки
END_VAR

(* ---- Fb1oo1DSAIMatchesTable.method.impl.st ---- *)
// AUTO-GENERATED by cemgen 1.0.0 — не редактировать: правьте матрицу и запустите
//   python -m cemgen generate <файл матрицы .csv или .xlsx>
// Матрица: SIS-V101-CEM, объект V-101, ревизия B от 2026-10-19, SHA-256 сетки df2ed4841a9453ca
coUnit.TEST('VoteTruth_Fb1oo1DSAI_MatchesTable');
stCfg.eArch := E_VoteArch.Vote1oo1;
stCfg.ePolicy := E_DegradePolicy.DegradeSafe;
stCfg.eInput := E_SisInputKind.Analog;
stCfg.xDiHealthy := TRUE;
stCfg.eLimitDir := E_LimitDir.High;
stCfg.rTripLimit_eu := 50.0;
stCfg.rHyst_eu := 0.0;
stCfg.rDiscrepancyMax_eu := 0.0;
stCfg.tDiscrepancyDelay := T#0S;
stCfg.tBypassMax := T#1H;
stCfg.uiMaxBypass := 0;
FOR uiRow := 0 TO 7 DO
    RowInputs(uiRow := uiRow, uiChannels := 1, xBypass := FALSE, stIn := stIn, stCmd := stCmd);
    fbVote(stIn := stIn, stCmd := stCmd, stCfg := stCfg, xBypassPermit := TRUE, uiCause := 1,
        itfTime := fbTime);
    RowInputs(uiRow := uiRow, uiChannels := 1, xBypass := TRUE, stIn := stIn, stCmd := stCmd);
    fbVote(stIn := stIn, stCmd := stCmd, stCfg := stCfg, xBypassPermit := TRUE, uiCause := 1,
        itfTime := fbTime);
    bAct := EncodeFb(xTrip := fbVote.xTrip, stSts := fbVote.stSts);
    bExp := GVL_VoteTruthTable.TT_FB_1OO1_DS_AI[uiRow];
    xMiss := bAct <> bExp;
    xFirst := xMiss AND uiMismatch = 0;
    uiFirstRow := SEL(xFirst, uiFirstRow, uiRow);
    bFirstExp := SEL(xFirst, bFirstExp, bExp);
    bFirstAct := SEL(xFirst, bFirstAct, bAct);
    uiMismatch := uiMismatch + BOOL_TO_UINT(xMiss);
END_FOR
AssertEquals_UINT(Expected := 0, Actual := uiMismatch,
    Message := MismatchText(sTable := 'TT_FB_1OO1_DS_AI', uiRow := uiFirstRow, bExpected := bFirstExp,
        bActual := bFirstAct));
coUnit.TEST_FINISHED();

(* ---- Fb1oo1DSDIMatchesTable.method.decl.st ---- *)
// AUTO-GENERATED by cemgen 1.0.0 — не редактировать: правьте матрицу и запустите
//   python -m cemgen generate <файл матрицы .csv или .xlsx>
// Матрица: SIS-V101-CEM, объект V-101, ревизия B от 2026-10-19, SHA-256 сетки df2ed4841a9453ca
// Назначение: тест VoteTruth_Fb1oo1DSDI_MatchesTable набора FB_VoteTruth_Test.
// Автор:      kr0nsch; код — генератор cemgen
// Версия:     1.0.0
// Документ:   docs/DESIGN.md, раздел «10. Генератор cemgen»; docs/cause_effect_matrix.md
// ВНИМАНИЕ:   код демонстрационный и не предназначен для систем безопасности. Реальная ПАЗ требует
//             определения SIL, сертифицированных аппаратных и программных средств и валидации по
//             ГОСТ Р МЭК 61511.
// FB_Voting, схема 1oo1, политика DegradeSafe, дискретные каналы: все 8 сочетаний «требование ×
// достоверность × запрос байпаса» совпадают с таблицей TT_FB_1OO1_DS_DI. На строку — два вызова одного
// экземпляра: без запросов байпаса (сброс байпасов прошлой строки) и с полной строкой.
METHOD PRIVATE Fb1oo1DSDIMatchesTable
VAR
    fbTime     : PL.FB_FakeTime;   // время не меняется
    fbVote     : FB_Voting;        // ФБ под тестом, один экземпляр на все строки
    stCfg      : ST_VotingCfg;     // конфигурация теста уровня 2
    stIn       : ST_VoteIn;        // входы строки
    stCmd      : ST_VoteCmd;       // запросы байпаса строки
    uiRow      : UINT;             // строка таблицы
    bAct       : BYTE;             // фактический байт результата
    bExp       : BYTE;             // ожидаемый байт из таблицы
    xMiss      : BOOL;             // строка не совпала
    xFirst     : BOOL;             // первая несовпавшая строка
    uiMismatch : UINT;             // несовпавших строк
    uiFirstRow : UINT;             // первая несовпавшая строка
    bFirstExp  : BYTE;             // ожидаемый байт первой несовпавшей строки
    bFirstAct  : BYTE;             // фактический байт первой несовпавшей строки
END_VAR

(* ---- Fb1oo1DSDIMatchesTable.method.impl.st ---- *)
// AUTO-GENERATED by cemgen 1.0.0 — не редактировать: правьте матрицу и запустите
//   python -m cemgen generate <файл матрицы .csv или .xlsx>
// Матрица: SIS-V101-CEM, объект V-101, ревизия B от 2026-10-19, SHA-256 сетки df2ed4841a9453ca
coUnit.TEST('VoteTruth_Fb1oo1DSDI_MatchesTable');
stCfg.eArch := E_VoteArch.Vote1oo1;
stCfg.ePolicy := E_DegradePolicy.DegradeSafe;
stCfg.eInput := E_SisInputKind.Discrete;
stCfg.xDiHealthy := TRUE;
stCfg.eLimitDir := E_LimitDir.High;
stCfg.rTripLimit_eu := 50.0;
stCfg.rHyst_eu := 0.0;
stCfg.rDiscrepancyMax_eu := 0.0;
stCfg.tDiscrepancyDelay := T#0S;
stCfg.tBypassMax := T#1H;
stCfg.uiMaxBypass := 0;
FOR uiRow := 0 TO 7 DO
    RowInputs(uiRow := uiRow, uiChannels := 1, xBypass := FALSE, stIn := stIn, stCmd := stCmd);
    fbVote(stIn := stIn, stCmd := stCmd, stCfg := stCfg, xBypassPermit := TRUE, uiCause := 1,
        itfTime := fbTime);
    RowInputs(uiRow := uiRow, uiChannels := 1, xBypass := TRUE, stIn := stIn, stCmd := stCmd);
    fbVote(stIn := stIn, stCmd := stCmd, stCfg := stCfg, xBypassPermit := TRUE, uiCause := 1,
        itfTime := fbTime);
    bAct := EncodeFb(xTrip := fbVote.xTrip, stSts := fbVote.stSts);
    bExp := GVL_VoteTruthTable.TT_FB_1OO1_DS_DI[uiRow];
    xMiss := bAct <> bExp;
    xFirst := xMiss AND uiMismatch = 0;
    uiFirstRow := SEL(xFirst, uiFirstRow, uiRow);
    bFirstExp := SEL(xFirst, bFirstExp, bExp);
    bFirstAct := SEL(xFirst, bFirstAct, bAct);
    uiMismatch := uiMismatch + BOOL_TO_UINT(xMiss);
END_FOR
AssertEquals_UINT(Expected := 0, Actual := uiMismatch,
    Message := MismatchText(sTable := 'TT_FB_1OO1_DS_DI', uiRow := uiFirstRow, bExpected := bFirstExp,
        bActual := bFirstAct));
coUnit.TEST_FINISHED();

(* ---- Fb1oo1VTAIMatchesTable.method.decl.st ---- *)
// AUTO-GENERATED by cemgen 1.0.0 — не редактировать: правьте матрицу и запустите
//   python -m cemgen generate <файл матрицы .csv или .xlsx>
// Матрица: SIS-V101-CEM, объект V-101, ревизия B от 2026-10-19, SHA-256 сетки df2ed4841a9453ca
// Назначение: тест VoteTruth_Fb1oo1VTAI_MatchesTable набора FB_VoteTruth_Test.
// Автор:      kr0nsch; код — генератор cemgen
// Версия:     1.0.0
// Документ:   docs/DESIGN.md, раздел «10. Генератор cemgen»; docs/cause_effect_matrix.md
// ВНИМАНИЕ:   код демонстрационный и не предназначен для систем безопасности. Реальная ПАЗ требует
//             определения SIL, сертифицированных аппаратных и программных средств и валидации по
//             ГОСТ Р МЭК 61511.
// FB_Voting, схема 1oo1, политика VoteTrip, аналоговые каналы: все 8 сочетаний «требование ×
// достоверность × запрос байпаса» совпадают с таблицей TT_FB_1OO1_VT_AI. На строку — два вызова одного
// экземпляра: без запросов байпаса (сброс байпасов прошлой строки) и с полной строкой.
METHOD PRIVATE Fb1oo1VTAIMatchesTable
VAR
    fbTime     : PL.FB_FakeTime;   // время не меняется
    fbVote     : FB_Voting;        // ФБ под тестом, один экземпляр на все строки
    stCfg      : ST_VotingCfg;     // конфигурация теста уровня 2
    stIn       : ST_VoteIn;        // входы строки
    stCmd      : ST_VoteCmd;       // запросы байпаса строки
    uiRow      : UINT;             // строка таблицы
    bAct       : BYTE;             // фактический байт результата
    bExp       : BYTE;             // ожидаемый байт из таблицы
    xMiss      : BOOL;             // строка не совпала
    xFirst     : BOOL;             // первая несовпавшая строка
    uiMismatch : UINT;             // несовпавших строк
    uiFirstRow : UINT;             // первая несовпавшая строка
    bFirstExp  : BYTE;             // ожидаемый байт первой несовпавшей строки
    bFirstAct  : BYTE;             // фактический байт первой несовпавшей строки
END_VAR

(* ---- Fb1oo1VTAIMatchesTable.method.impl.st ---- *)
// AUTO-GENERATED by cemgen 1.0.0 — не редактировать: правьте матрицу и запустите
//   python -m cemgen generate <файл матрицы .csv или .xlsx>
// Матрица: SIS-V101-CEM, объект V-101, ревизия B от 2026-10-19, SHA-256 сетки df2ed4841a9453ca
coUnit.TEST('VoteTruth_Fb1oo1VTAI_MatchesTable');
stCfg.eArch := E_VoteArch.Vote1oo1;
stCfg.ePolicy := E_DegradePolicy.VoteTrip;
stCfg.eInput := E_SisInputKind.Analog;
stCfg.xDiHealthy := TRUE;
stCfg.eLimitDir := E_LimitDir.High;
stCfg.rTripLimit_eu := 50.0;
stCfg.rHyst_eu := 0.0;
stCfg.rDiscrepancyMax_eu := 0.0;
stCfg.tDiscrepancyDelay := T#0S;
stCfg.tBypassMax := T#1H;
stCfg.uiMaxBypass := 0;
FOR uiRow := 0 TO 7 DO
    RowInputs(uiRow := uiRow, uiChannels := 1, xBypass := FALSE, stIn := stIn, stCmd := stCmd);
    fbVote(stIn := stIn, stCmd := stCmd, stCfg := stCfg, xBypassPermit := TRUE, uiCause := 1,
        itfTime := fbTime);
    RowInputs(uiRow := uiRow, uiChannels := 1, xBypass := TRUE, stIn := stIn, stCmd := stCmd);
    fbVote(stIn := stIn, stCmd := stCmd, stCfg := stCfg, xBypassPermit := TRUE, uiCause := 1,
        itfTime := fbTime);
    bAct := EncodeFb(xTrip := fbVote.xTrip, stSts := fbVote.stSts);
    bExp := GVL_VoteTruthTable.TT_FB_1OO1_VT_AI[uiRow];
    xMiss := bAct <> bExp;
    xFirst := xMiss AND uiMismatch = 0;
    uiFirstRow := SEL(xFirst, uiFirstRow, uiRow);
    bFirstExp := SEL(xFirst, bFirstExp, bExp);
    bFirstAct := SEL(xFirst, bFirstAct, bAct);
    uiMismatch := uiMismatch + BOOL_TO_UINT(xMiss);
END_FOR
AssertEquals_UINT(Expected := 0, Actual := uiMismatch,
    Message := MismatchText(sTable := 'TT_FB_1OO1_VT_AI', uiRow := uiFirstRow, bExpected := bFirstExp,
        bActual := bFirstAct));
coUnit.TEST_FINISHED();

(* ---- Fb1oo1VTDIMatchesTable.method.decl.st ---- *)
// AUTO-GENERATED by cemgen 1.0.0 — не редактировать: правьте матрицу и запустите
//   python -m cemgen generate <файл матрицы .csv или .xlsx>
// Матрица: SIS-V101-CEM, объект V-101, ревизия B от 2026-10-19, SHA-256 сетки df2ed4841a9453ca
// Назначение: тест VoteTruth_Fb1oo1VTDI_MatchesTable набора FB_VoteTruth_Test.
// Автор:      kr0nsch; код — генератор cemgen
// Версия:     1.0.0
// Документ:   docs/DESIGN.md, раздел «10. Генератор cemgen»; docs/cause_effect_matrix.md
// ВНИМАНИЕ:   код демонстрационный и не предназначен для систем безопасности. Реальная ПАЗ требует
//             определения SIL, сертифицированных аппаратных и программных средств и валидации по
//             ГОСТ Р МЭК 61511.
// FB_Voting, схема 1oo1, политика VoteTrip, дискретные каналы: все 8 сочетаний «требование ×
// достоверность × запрос байпаса» совпадают с таблицей TT_FB_1OO1_VT_DI. На строку — два вызова одного
// экземпляра: без запросов байпаса (сброс байпасов прошлой строки) и с полной строкой.
METHOD PRIVATE Fb1oo1VTDIMatchesTable
VAR
    fbTime     : PL.FB_FakeTime;   // время не меняется
    fbVote     : FB_Voting;        // ФБ под тестом, один экземпляр на все строки
    stCfg      : ST_VotingCfg;     // конфигурация теста уровня 2
    stIn       : ST_VoteIn;        // входы строки
    stCmd      : ST_VoteCmd;       // запросы байпаса строки
    uiRow      : UINT;             // строка таблицы
    bAct       : BYTE;             // фактический байт результата
    bExp       : BYTE;             // ожидаемый байт из таблицы
    xMiss      : BOOL;             // строка не совпала
    xFirst     : BOOL;             // первая несовпавшая строка
    uiMismatch : UINT;             // несовпавших строк
    uiFirstRow : UINT;             // первая несовпавшая строка
    bFirstExp  : BYTE;             // ожидаемый байт первой несовпавшей строки
    bFirstAct  : BYTE;             // фактический байт первой несовпавшей строки
END_VAR

(* ---- Fb1oo1VTDIMatchesTable.method.impl.st ---- *)
// AUTO-GENERATED by cemgen 1.0.0 — не редактировать: правьте матрицу и запустите
//   python -m cemgen generate <файл матрицы .csv или .xlsx>
// Матрица: SIS-V101-CEM, объект V-101, ревизия B от 2026-10-19, SHA-256 сетки df2ed4841a9453ca
coUnit.TEST('VoteTruth_Fb1oo1VTDI_MatchesTable');
stCfg.eArch := E_VoteArch.Vote1oo1;
stCfg.ePolicy := E_DegradePolicy.VoteTrip;
stCfg.eInput := E_SisInputKind.Discrete;
stCfg.xDiHealthy := TRUE;
stCfg.eLimitDir := E_LimitDir.High;
stCfg.rTripLimit_eu := 50.0;
stCfg.rHyst_eu := 0.0;
stCfg.rDiscrepancyMax_eu := 0.0;
stCfg.tDiscrepancyDelay := T#0S;
stCfg.tBypassMax := T#1H;
stCfg.uiMaxBypass := 0;
FOR uiRow := 0 TO 7 DO
    RowInputs(uiRow := uiRow, uiChannels := 1, xBypass := FALSE, stIn := stIn, stCmd := stCmd);
    fbVote(stIn := stIn, stCmd := stCmd, stCfg := stCfg, xBypassPermit := TRUE, uiCause := 1,
        itfTime := fbTime);
    RowInputs(uiRow := uiRow, uiChannels := 1, xBypass := TRUE, stIn := stIn, stCmd := stCmd);
    fbVote(stIn := stIn, stCmd := stCmd, stCfg := stCfg, xBypassPermit := TRUE, uiCause := 1,
        itfTime := fbTime);
    bAct := EncodeFb(xTrip := fbVote.xTrip, stSts := fbVote.stSts);
    bExp := GVL_VoteTruthTable.TT_FB_1OO1_VT_DI[uiRow];
    xMiss := bAct <> bExp;
    xFirst := xMiss AND uiMismatch = 0;
    uiFirstRow := SEL(xFirst, uiFirstRow, uiRow);
    bFirstExp := SEL(xFirst, bFirstExp, bExp);
    bFirstAct := SEL(xFirst, bFirstAct, bAct);
    uiMismatch := uiMismatch + BOOL_TO_UINT(xMiss);
END_FOR
AssertEquals_UINT(Expected := 0, Actual := uiMismatch,
    Message := MismatchText(sTable := 'TT_FB_1OO1_VT_DI', uiRow := uiFirstRow, bExpected := bFirstExp,
        bActual := bFirstAct));
coUnit.TEST_FINISHED();

(* ---- Fb1oo2DAAIMatchesTable.method.decl.st ---- *)
// AUTO-GENERATED by cemgen 1.0.0 — не редактировать: правьте матрицу и запустите
//   python -m cemgen generate <файл матрицы .csv или .xlsx>
// Матрица: SIS-V101-CEM, объект V-101, ревизия B от 2026-10-19, SHA-256 сетки df2ed4841a9453ca
// Назначение: тест VoteTruth_Fb1oo2DAAI_MatchesTable набора FB_VoteTruth_Test.
// Автор:      kr0nsch; код — генератор cemgen
// Версия:     1.0.0
// Документ:   docs/DESIGN.md, раздел «10. Генератор cemgen»; docs/cause_effect_matrix.md
// ВНИМАНИЕ:   код демонстрационный и не предназначен для систем безопасности. Реальная ПАЗ требует
//             определения SIL, сертифицированных аппаратных и программных средств и валидации по
//             ГОСТ Р МЭК 61511.
// FB_Voting, схема 1oo2, политика DegradeAvailable, аналоговые каналы: все 64 сочетаний «требование ×
// достоверность × запрос байпаса» совпадают с таблицей TT_FB_1OO2_DA_AI. На строку — два вызова одного
// экземпляра: без запросов байпаса (сброс байпасов прошлой строки) и с полной строкой.
METHOD PRIVATE Fb1oo2DAAIMatchesTable
VAR
    fbTime     : PL.FB_FakeTime;   // время не меняется
    fbVote     : FB_Voting;        // ФБ под тестом, один экземпляр на все строки
    stCfg      : ST_VotingCfg;     // конфигурация теста уровня 2
    stIn       : ST_VoteIn;        // входы строки
    stCmd      : ST_VoteCmd;       // запросы байпаса строки
    uiRow      : UINT;             // строка таблицы
    bAct       : BYTE;             // фактический байт результата
    bExp       : BYTE;             // ожидаемый байт из таблицы
    xMiss      : BOOL;             // строка не совпала
    xFirst     : BOOL;             // первая несовпавшая строка
    uiMismatch : UINT;             // несовпавших строк
    uiFirstRow : UINT;             // первая несовпавшая строка
    bFirstExp  : BYTE;             // ожидаемый байт первой несовпавшей строки
    bFirstAct  : BYTE;             // фактический байт первой несовпавшей строки
END_VAR

(* ---- Fb1oo2DAAIMatchesTable.method.impl.st ---- *)
// AUTO-GENERATED by cemgen 1.0.0 — не редактировать: правьте матрицу и запустите
//   python -m cemgen generate <файл матрицы .csv или .xlsx>
// Матрица: SIS-V101-CEM, объект V-101, ревизия B от 2026-10-19, SHA-256 сетки df2ed4841a9453ca
coUnit.TEST('VoteTruth_Fb1oo2DAAI_MatchesTable');
stCfg.eArch := E_VoteArch.Vote1oo2;
stCfg.ePolicy := E_DegradePolicy.DegradeAvailable;
stCfg.eInput := E_SisInputKind.Analog;
stCfg.xDiHealthy := TRUE;
stCfg.eLimitDir := E_LimitDir.High;
stCfg.rTripLimit_eu := 50.0;
stCfg.rHyst_eu := 0.0;
stCfg.rDiscrepancyMax_eu := 0.0;
stCfg.tDiscrepancyDelay := T#0S;
stCfg.tBypassMax := T#1H;
stCfg.uiMaxBypass := 1;
FOR uiRow := 0 TO 63 DO
    RowInputs(uiRow := uiRow, uiChannels := 2, xBypass := FALSE, stIn := stIn, stCmd := stCmd);
    fbVote(stIn := stIn, stCmd := stCmd, stCfg := stCfg, xBypassPermit := TRUE, uiCause := 1,
        itfTime := fbTime);
    RowInputs(uiRow := uiRow, uiChannels := 2, xBypass := TRUE, stIn := stIn, stCmd := stCmd);
    fbVote(stIn := stIn, stCmd := stCmd, stCfg := stCfg, xBypassPermit := TRUE, uiCause := 1,
        itfTime := fbTime);
    bAct := EncodeFb(xTrip := fbVote.xTrip, stSts := fbVote.stSts);
    bExp := GVL_VoteTruthTable.TT_FB_1OO2_DA_AI[uiRow];
    xMiss := bAct <> bExp;
    xFirst := xMiss AND uiMismatch = 0;
    uiFirstRow := SEL(xFirst, uiFirstRow, uiRow);
    bFirstExp := SEL(xFirst, bFirstExp, bExp);
    bFirstAct := SEL(xFirst, bFirstAct, bAct);
    uiMismatch := uiMismatch + BOOL_TO_UINT(xMiss);
END_FOR
AssertEquals_UINT(Expected := 0, Actual := uiMismatch,
    Message := MismatchText(sTable := 'TT_FB_1OO2_DA_AI', uiRow := uiFirstRow, bExpected := bFirstExp,
        bActual := bFirstAct));
coUnit.TEST_FINISHED();

(* ---- Fb1oo2DADIMatchesTable.method.decl.st ---- *)
// AUTO-GENERATED by cemgen 1.0.0 — не редактировать: правьте матрицу и запустите
//   python -m cemgen generate <файл матрицы .csv или .xlsx>
// Матрица: SIS-V101-CEM, объект V-101, ревизия B от 2026-10-19, SHA-256 сетки df2ed4841a9453ca
// Назначение: тест VoteTruth_Fb1oo2DADI_MatchesTable набора FB_VoteTruth_Test.
// Автор:      kr0nsch; код — генератор cemgen
// Версия:     1.0.0
// Документ:   docs/DESIGN.md, раздел «10. Генератор cemgen»; docs/cause_effect_matrix.md
// ВНИМАНИЕ:   код демонстрационный и не предназначен для систем безопасности. Реальная ПАЗ требует
//             определения SIL, сертифицированных аппаратных и программных средств и валидации по
//             ГОСТ Р МЭК 61511.
// FB_Voting, схема 1oo2, политика DegradeAvailable, дискретные каналы: все 64 сочетаний «требование ×
// достоверность × запрос байпаса» совпадают с таблицей TT_FB_1OO2_DA_DI. На строку — два вызова одного
// экземпляра: без запросов байпаса (сброс байпасов прошлой строки) и с полной строкой.
METHOD PRIVATE Fb1oo2DADIMatchesTable
VAR
    fbTime     : PL.FB_FakeTime;   // время не меняется
    fbVote     : FB_Voting;        // ФБ под тестом, один экземпляр на все строки
    stCfg      : ST_VotingCfg;     // конфигурация теста уровня 2
    stIn       : ST_VoteIn;        // входы строки
    stCmd      : ST_VoteCmd;       // запросы байпаса строки
    uiRow      : UINT;             // строка таблицы
    bAct       : BYTE;             // фактический байт результата
    bExp       : BYTE;             // ожидаемый байт из таблицы
    xMiss      : BOOL;             // строка не совпала
    xFirst     : BOOL;             // первая несовпавшая строка
    uiMismatch : UINT;             // несовпавших строк
    uiFirstRow : UINT;             // первая несовпавшая строка
    bFirstExp  : BYTE;             // ожидаемый байт первой несовпавшей строки
    bFirstAct  : BYTE;             // фактический байт первой несовпавшей строки
END_VAR

(* ---- Fb1oo2DADIMatchesTable.method.impl.st ---- *)
// AUTO-GENERATED by cemgen 1.0.0 — не редактировать: правьте матрицу и запустите
//   python -m cemgen generate <файл матрицы .csv или .xlsx>
// Матрица: SIS-V101-CEM, объект V-101, ревизия B от 2026-10-19, SHA-256 сетки df2ed4841a9453ca
coUnit.TEST('VoteTruth_Fb1oo2DADI_MatchesTable');
stCfg.eArch := E_VoteArch.Vote1oo2;
stCfg.ePolicy := E_DegradePolicy.DegradeAvailable;
stCfg.eInput := E_SisInputKind.Discrete;
stCfg.xDiHealthy := TRUE;
stCfg.eLimitDir := E_LimitDir.High;
stCfg.rTripLimit_eu := 50.0;
stCfg.rHyst_eu := 0.0;
stCfg.rDiscrepancyMax_eu := 0.0;
stCfg.tDiscrepancyDelay := T#0S;
stCfg.tBypassMax := T#1H;
stCfg.uiMaxBypass := 1;
FOR uiRow := 0 TO 63 DO
    RowInputs(uiRow := uiRow, uiChannels := 2, xBypass := FALSE, stIn := stIn, stCmd := stCmd);
    fbVote(stIn := stIn, stCmd := stCmd, stCfg := stCfg, xBypassPermit := TRUE, uiCause := 1,
        itfTime := fbTime);
    RowInputs(uiRow := uiRow, uiChannels := 2, xBypass := TRUE, stIn := stIn, stCmd := stCmd);
    fbVote(stIn := stIn, stCmd := stCmd, stCfg := stCfg, xBypassPermit := TRUE, uiCause := 1,
        itfTime := fbTime);
    bAct := EncodeFb(xTrip := fbVote.xTrip, stSts := fbVote.stSts);
    bExp := GVL_VoteTruthTable.TT_FB_1OO2_DA_DI[uiRow];
    xMiss := bAct <> bExp;
    xFirst := xMiss AND uiMismatch = 0;
    uiFirstRow := SEL(xFirst, uiFirstRow, uiRow);
    bFirstExp := SEL(xFirst, bFirstExp, bExp);
    bFirstAct := SEL(xFirst, bFirstAct, bAct);
    uiMismatch := uiMismatch + BOOL_TO_UINT(xMiss);
END_FOR
AssertEquals_UINT(Expected := 0, Actual := uiMismatch,
    Message := MismatchText(sTable := 'TT_FB_1OO2_DA_DI', uiRow := uiFirstRow, bExpected := bFirstExp,
        bActual := bFirstAct));
coUnit.TEST_FINISHED();

(* ---- Fb1oo2DSAIMatchesTable.method.decl.st ---- *)
// AUTO-GENERATED by cemgen 1.0.0 — не редактировать: правьте матрицу и запустите
//   python -m cemgen generate <файл матрицы .csv или .xlsx>
// Матрица: SIS-V101-CEM, объект V-101, ревизия B от 2026-10-19, SHA-256 сетки df2ed4841a9453ca
// Назначение: тест VoteTruth_Fb1oo2DSAI_MatchesTable набора FB_VoteTruth_Test.
// Автор:      kr0nsch; код — генератор cemgen
// Версия:     1.0.0
// Документ:   docs/DESIGN.md, раздел «10. Генератор cemgen»; docs/cause_effect_matrix.md
// ВНИМАНИЕ:   код демонстрационный и не предназначен для систем безопасности. Реальная ПАЗ требует
//             определения SIL, сертифицированных аппаратных и программных средств и валидации по
//             ГОСТ Р МЭК 61511.
// FB_Voting, схема 1oo2, политика DegradeSafe, аналоговые каналы: все 64 сочетаний «требование ×
// достоверность × запрос байпаса» совпадают с таблицей TT_FB_1OO2_DS_AI. На строку — два вызова одного
// экземпляра: без запросов байпаса (сброс байпасов прошлой строки) и с полной строкой.
METHOD PRIVATE Fb1oo2DSAIMatchesTable
VAR
    fbTime     : PL.FB_FakeTime;   // время не меняется
    fbVote     : FB_Voting;        // ФБ под тестом, один экземпляр на все строки
    stCfg      : ST_VotingCfg;     // конфигурация теста уровня 2
    stIn       : ST_VoteIn;        // входы строки
    stCmd      : ST_VoteCmd;       // запросы байпаса строки
    uiRow      : UINT;             // строка таблицы
    bAct       : BYTE;             // фактический байт результата
    bExp       : BYTE;             // ожидаемый байт из таблицы
    xMiss      : BOOL;             // строка не совпала
    xFirst     : BOOL;             // первая несовпавшая строка
    uiMismatch : UINT;             // несовпавших строк
    uiFirstRow : UINT;             // первая несовпавшая строка
    bFirstExp  : BYTE;             // ожидаемый байт первой несовпавшей строки
    bFirstAct  : BYTE;             // фактический байт первой несовпавшей строки
END_VAR

(* ---- Fb1oo2DSAIMatchesTable.method.impl.st ---- *)
// AUTO-GENERATED by cemgen 1.0.0 — не редактировать: правьте матрицу и запустите
//   python -m cemgen generate <файл матрицы .csv или .xlsx>
// Матрица: SIS-V101-CEM, объект V-101, ревизия B от 2026-10-19, SHA-256 сетки df2ed4841a9453ca
coUnit.TEST('VoteTruth_Fb1oo2DSAI_MatchesTable');
stCfg.eArch := E_VoteArch.Vote1oo2;
stCfg.ePolicy := E_DegradePolicy.DegradeSafe;
stCfg.eInput := E_SisInputKind.Analog;
stCfg.xDiHealthy := TRUE;
stCfg.eLimitDir := E_LimitDir.High;
stCfg.rTripLimit_eu := 50.0;
stCfg.rHyst_eu := 0.0;
stCfg.rDiscrepancyMax_eu := 0.0;
stCfg.tDiscrepancyDelay := T#0S;
stCfg.tBypassMax := T#1H;
stCfg.uiMaxBypass := 1;
FOR uiRow := 0 TO 63 DO
    RowInputs(uiRow := uiRow, uiChannels := 2, xBypass := FALSE, stIn := stIn, stCmd := stCmd);
    fbVote(stIn := stIn, stCmd := stCmd, stCfg := stCfg, xBypassPermit := TRUE, uiCause := 1,
        itfTime := fbTime);
    RowInputs(uiRow := uiRow, uiChannels := 2, xBypass := TRUE, stIn := stIn, stCmd := stCmd);
    fbVote(stIn := stIn, stCmd := stCmd, stCfg := stCfg, xBypassPermit := TRUE, uiCause := 1,
        itfTime := fbTime);
    bAct := EncodeFb(xTrip := fbVote.xTrip, stSts := fbVote.stSts);
    bExp := GVL_VoteTruthTable.TT_FB_1OO2_DS_AI[uiRow];
    xMiss := bAct <> bExp;
    xFirst := xMiss AND uiMismatch = 0;
    uiFirstRow := SEL(xFirst, uiFirstRow, uiRow);
    bFirstExp := SEL(xFirst, bFirstExp, bExp);
    bFirstAct := SEL(xFirst, bFirstAct, bAct);
    uiMismatch := uiMismatch + BOOL_TO_UINT(xMiss);
END_FOR
AssertEquals_UINT(Expected := 0, Actual := uiMismatch,
    Message := MismatchText(sTable := 'TT_FB_1OO2_DS_AI', uiRow := uiFirstRow, bExpected := bFirstExp,
        bActual := bFirstAct));
coUnit.TEST_FINISHED();

(* ---- Fb1oo2DSDIMatchesTable.method.decl.st ---- *)
// AUTO-GENERATED by cemgen 1.0.0 — не редактировать: правьте матрицу и запустите
//   python -m cemgen generate <файл матрицы .csv или .xlsx>
// Матрица: SIS-V101-CEM, объект V-101, ревизия B от 2026-10-19, SHA-256 сетки df2ed4841a9453ca
// Назначение: тест VoteTruth_Fb1oo2DSDI_MatchesTable набора FB_VoteTruth_Test.
// Автор:      kr0nsch; код — генератор cemgen
// Версия:     1.0.0
// Документ:   docs/DESIGN.md, раздел «10. Генератор cemgen»; docs/cause_effect_matrix.md
// ВНИМАНИЕ:   код демонстрационный и не предназначен для систем безопасности. Реальная ПАЗ требует
//             определения SIL, сертифицированных аппаратных и программных средств и валидации по
//             ГОСТ Р МЭК 61511.
// FB_Voting, схема 1oo2, политика DegradeSafe, дискретные каналы: все 64 сочетаний «требование ×
// достоверность × запрос байпаса» совпадают с таблицей TT_FB_1OO2_DS_DI. На строку — два вызова одного
// экземпляра: без запросов байпаса (сброс байпасов прошлой строки) и с полной строкой.
METHOD PRIVATE Fb1oo2DSDIMatchesTable
VAR
    fbTime     : PL.FB_FakeTime;   // время не меняется
    fbVote     : FB_Voting;        // ФБ под тестом, один экземпляр на все строки
    stCfg      : ST_VotingCfg;     // конфигурация теста уровня 2
    stIn       : ST_VoteIn;        // входы строки
    stCmd      : ST_VoteCmd;       // запросы байпаса строки
    uiRow      : UINT;             // строка таблицы
    bAct       : BYTE;             // фактический байт результата
    bExp       : BYTE;             // ожидаемый байт из таблицы
    xMiss      : BOOL;             // строка не совпала
    xFirst     : BOOL;             // первая несовпавшая строка
    uiMismatch : UINT;             // несовпавших строк
    uiFirstRow : UINT;             // первая несовпавшая строка
    bFirstExp  : BYTE;             // ожидаемый байт первой несовпавшей строки
    bFirstAct  : BYTE;             // фактический байт первой несовпавшей строки
END_VAR

(* ---- Fb1oo2DSDIMatchesTable.method.impl.st ---- *)
// AUTO-GENERATED by cemgen 1.0.0 — не редактировать: правьте матрицу и запустите
//   python -m cemgen generate <файл матрицы .csv или .xlsx>
// Матрица: SIS-V101-CEM, объект V-101, ревизия B от 2026-10-19, SHA-256 сетки df2ed4841a9453ca
coUnit.TEST('VoteTruth_Fb1oo2DSDI_MatchesTable');
stCfg.eArch := E_VoteArch.Vote1oo2;
stCfg.ePolicy := E_DegradePolicy.DegradeSafe;
stCfg.eInput := E_SisInputKind.Discrete;
stCfg.xDiHealthy := TRUE;
stCfg.eLimitDir := E_LimitDir.High;
stCfg.rTripLimit_eu := 50.0;
stCfg.rHyst_eu := 0.0;
stCfg.rDiscrepancyMax_eu := 0.0;
stCfg.tDiscrepancyDelay := T#0S;
stCfg.tBypassMax := T#1H;
stCfg.uiMaxBypass := 1;
FOR uiRow := 0 TO 63 DO
    RowInputs(uiRow := uiRow, uiChannels := 2, xBypass := FALSE, stIn := stIn, stCmd := stCmd);
    fbVote(stIn := stIn, stCmd := stCmd, stCfg := stCfg, xBypassPermit := TRUE, uiCause := 1,
        itfTime := fbTime);
    RowInputs(uiRow := uiRow, uiChannels := 2, xBypass := TRUE, stIn := stIn, stCmd := stCmd);
    fbVote(stIn := stIn, stCmd := stCmd, stCfg := stCfg, xBypassPermit := TRUE, uiCause := 1,
        itfTime := fbTime);
    bAct := EncodeFb(xTrip := fbVote.xTrip, stSts := fbVote.stSts);
    bExp := GVL_VoteTruthTable.TT_FB_1OO2_DS_DI[uiRow];
    xMiss := bAct <> bExp;
    xFirst := xMiss AND uiMismatch = 0;
    uiFirstRow := SEL(xFirst, uiFirstRow, uiRow);
    bFirstExp := SEL(xFirst, bFirstExp, bExp);
    bFirstAct := SEL(xFirst, bFirstAct, bAct);
    uiMismatch := uiMismatch + BOOL_TO_UINT(xMiss);
END_FOR
AssertEquals_UINT(Expected := 0, Actual := uiMismatch,
    Message := MismatchText(sTable := 'TT_FB_1OO2_DS_DI', uiRow := uiFirstRow, bExpected := bFirstExp,
        bActual := bFirstAct));
coUnit.TEST_FINISHED();

(* ---- Fb1oo2VTAIMatchesTable.method.decl.st ---- *)
// AUTO-GENERATED by cemgen 1.0.0 — не редактировать: правьте матрицу и запустите
//   python -m cemgen generate <файл матрицы .csv или .xlsx>
// Матрица: SIS-V101-CEM, объект V-101, ревизия B от 2026-10-19, SHA-256 сетки df2ed4841a9453ca
// Назначение: тест VoteTruth_Fb1oo2VTAI_MatchesTable набора FB_VoteTruth_Test.
// Автор:      kr0nsch; код — генератор cemgen
// Версия:     1.0.0
// Документ:   docs/DESIGN.md, раздел «10. Генератор cemgen»; docs/cause_effect_matrix.md
// ВНИМАНИЕ:   код демонстрационный и не предназначен для систем безопасности. Реальная ПАЗ требует
//             определения SIL, сертифицированных аппаратных и программных средств и валидации по
//             ГОСТ Р МЭК 61511.
// FB_Voting, схема 1oo2, политика VoteTrip, аналоговые каналы: все 64 сочетаний «требование ×
// достоверность × запрос байпаса» совпадают с таблицей TT_FB_1OO2_VT_AI. На строку — два вызова одного
// экземпляра: без запросов байпаса (сброс байпасов прошлой строки) и с полной строкой.
METHOD PRIVATE Fb1oo2VTAIMatchesTable
VAR
    fbTime     : PL.FB_FakeTime;   // время не меняется
    fbVote     : FB_Voting;        // ФБ под тестом, один экземпляр на все строки
    stCfg      : ST_VotingCfg;     // конфигурация теста уровня 2
    stIn       : ST_VoteIn;        // входы строки
    stCmd      : ST_VoteCmd;       // запросы байпаса строки
    uiRow      : UINT;             // строка таблицы
    bAct       : BYTE;             // фактический байт результата
    bExp       : BYTE;             // ожидаемый байт из таблицы
    xMiss      : BOOL;             // строка не совпала
    xFirst     : BOOL;             // первая несовпавшая строка
    uiMismatch : UINT;             // несовпавших строк
    uiFirstRow : UINT;             // первая несовпавшая строка
    bFirstExp  : BYTE;             // ожидаемый байт первой несовпавшей строки
    bFirstAct  : BYTE;             // фактический байт первой несовпавшей строки
END_VAR

(* ---- Fb1oo2VTAIMatchesTable.method.impl.st ---- *)
// AUTO-GENERATED by cemgen 1.0.0 — не редактировать: правьте матрицу и запустите
//   python -m cemgen generate <файл матрицы .csv или .xlsx>
// Матрица: SIS-V101-CEM, объект V-101, ревизия B от 2026-10-19, SHA-256 сетки df2ed4841a9453ca
coUnit.TEST('VoteTruth_Fb1oo2VTAI_MatchesTable');
stCfg.eArch := E_VoteArch.Vote1oo2;
stCfg.ePolicy := E_DegradePolicy.VoteTrip;
stCfg.eInput := E_SisInputKind.Analog;
stCfg.xDiHealthy := TRUE;
stCfg.eLimitDir := E_LimitDir.High;
stCfg.rTripLimit_eu := 50.0;
stCfg.rHyst_eu := 0.0;
stCfg.rDiscrepancyMax_eu := 0.0;
stCfg.tDiscrepancyDelay := T#0S;
stCfg.tBypassMax := T#1H;
stCfg.uiMaxBypass := 1;
FOR uiRow := 0 TO 63 DO
    RowInputs(uiRow := uiRow, uiChannels := 2, xBypass := FALSE, stIn := stIn, stCmd := stCmd);
    fbVote(stIn := stIn, stCmd := stCmd, stCfg := stCfg, xBypassPermit := TRUE, uiCause := 1,
        itfTime := fbTime);
    RowInputs(uiRow := uiRow, uiChannels := 2, xBypass := TRUE, stIn := stIn, stCmd := stCmd);
    fbVote(stIn := stIn, stCmd := stCmd, stCfg := stCfg, xBypassPermit := TRUE, uiCause := 1,
        itfTime := fbTime);
    bAct := EncodeFb(xTrip := fbVote.xTrip, stSts := fbVote.stSts);
    bExp := GVL_VoteTruthTable.TT_FB_1OO2_VT_AI[uiRow];
    xMiss := bAct <> bExp;
    xFirst := xMiss AND uiMismatch = 0;
    uiFirstRow := SEL(xFirst, uiFirstRow, uiRow);
    bFirstExp := SEL(xFirst, bFirstExp, bExp);
    bFirstAct := SEL(xFirst, bFirstAct, bAct);
    uiMismatch := uiMismatch + BOOL_TO_UINT(xMiss);
END_FOR
AssertEquals_UINT(Expected := 0, Actual := uiMismatch,
    Message := MismatchText(sTable := 'TT_FB_1OO2_VT_AI', uiRow := uiFirstRow, bExpected := bFirstExp,
        bActual := bFirstAct));
coUnit.TEST_FINISHED();

(* ---- Fb1oo2VTDIMatchesTable.method.decl.st ---- *)
// AUTO-GENERATED by cemgen 1.0.0 — не редактировать: правьте матрицу и запустите
//   python -m cemgen generate <файл матрицы .csv или .xlsx>
// Матрица: SIS-V101-CEM, объект V-101, ревизия B от 2026-10-19, SHA-256 сетки df2ed4841a9453ca
// Назначение: тест VoteTruth_Fb1oo2VTDI_MatchesTable набора FB_VoteTruth_Test.
// Автор:      kr0nsch; код — генератор cemgen
// Версия:     1.0.0
// Документ:   docs/DESIGN.md, раздел «10. Генератор cemgen»; docs/cause_effect_matrix.md
// ВНИМАНИЕ:   код демонстрационный и не предназначен для систем безопасности. Реальная ПАЗ требует
//             определения SIL, сертифицированных аппаратных и программных средств и валидации по
//             ГОСТ Р МЭК 61511.
// FB_Voting, схема 1oo2, политика VoteTrip, дискретные каналы: все 64 сочетаний «требование ×
// достоверность × запрос байпаса» совпадают с таблицей TT_FB_1OO2_VT_DI. На строку — два вызова одного
// экземпляра: без запросов байпаса (сброс байпасов прошлой строки) и с полной строкой.
METHOD PRIVATE Fb1oo2VTDIMatchesTable
VAR
    fbTime     : PL.FB_FakeTime;   // время не меняется
    fbVote     : FB_Voting;        // ФБ под тестом, один экземпляр на все строки
    stCfg      : ST_VotingCfg;     // конфигурация теста уровня 2
    stIn       : ST_VoteIn;        // входы строки
    stCmd      : ST_VoteCmd;       // запросы байпаса строки
    uiRow      : UINT;             // строка таблицы
    bAct       : BYTE;             // фактический байт результата
    bExp       : BYTE;             // ожидаемый байт из таблицы
    xMiss      : BOOL;             // строка не совпала
    xFirst     : BOOL;             // первая несовпавшая строка
    uiMismatch : UINT;             // несовпавших строк
    uiFirstRow : UINT;             // первая несовпавшая строка
    bFirstExp  : BYTE;             // ожидаемый байт первой несовпавшей строки
    bFirstAct  : BYTE;             // фактический байт первой несовпавшей строки
END_VAR

(* ---- Fb1oo2VTDIMatchesTable.method.impl.st ---- *)
// AUTO-GENERATED by cemgen 1.0.0 — не редактировать: правьте матрицу и запустите
//   python -m cemgen generate <файл матрицы .csv или .xlsx>
// Матрица: SIS-V101-CEM, объект V-101, ревизия B от 2026-10-19, SHA-256 сетки df2ed4841a9453ca
coUnit.TEST('VoteTruth_Fb1oo2VTDI_MatchesTable');
stCfg.eArch := E_VoteArch.Vote1oo2;
stCfg.ePolicy := E_DegradePolicy.VoteTrip;
stCfg.eInput := E_SisInputKind.Discrete;
stCfg.xDiHealthy := TRUE;
stCfg.eLimitDir := E_LimitDir.High;
stCfg.rTripLimit_eu := 50.0;
stCfg.rHyst_eu := 0.0;
stCfg.rDiscrepancyMax_eu := 0.0;
stCfg.tDiscrepancyDelay := T#0S;
stCfg.tBypassMax := T#1H;
stCfg.uiMaxBypass := 1;
FOR uiRow := 0 TO 63 DO
    RowInputs(uiRow := uiRow, uiChannels := 2, xBypass := FALSE, stIn := stIn, stCmd := stCmd);
    fbVote(stIn := stIn, stCmd := stCmd, stCfg := stCfg, xBypassPermit := TRUE, uiCause := 1,
        itfTime := fbTime);
    RowInputs(uiRow := uiRow, uiChannels := 2, xBypass := TRUE, stIn := stIn, stCmd := stCmd);
    fbVote(stIn := stIn, stCmd := stCmd, stCfg := stCfg, xBypassPermit := TRUE, uiCause := 1,
        itfTime := fbTime);
    bAct := EncodeFb(xTrip := fbVote.xTrip, stSts := fbVote.stSts);
    bExp := GVL_VoteTruthTable.TT_FB_1OO2_VT_DI[uiRow];
    xMiss := bAct <> bExp;
    xFirst := xMiss AND uiMismatch = 0;
    uiFirstRow := SEL(xFirst, uiFirstRow, uiRow);
    bFirstExp := SEL(xFirst, bFirstExp, bExp);
    bFirstAct := SEL(xFirst, bFirstAct, bAct);
    uiMismatch := uiMismatch + BOOL_TO_UINT(xMiss);
END_FOR
AssertEquals_UINT(Expected := 0, Actual := uiMismatch,
    Message := MismatchText(sTable := 'TT_FB_1OO2_VT_DI', uiRow := uiFirstRow, bExpected := bFirstExp,
        bActual := bFirstAct));
coUnit.TEST_FINISHED();

(* ---- Fb2oo2DAAIMatchesTable.method.decl.st ---- *)
// AUTO-GENERATED by cemgen 1.0.0 — не редактировать: правьте матрицу и запустите
//   python -m cemgen generate <файл матрицы .csv или .xlsx>
// Матрица: SIS-V101-CEM, объект V-101, ревизия B от 2026-10-19, SHA-256 сетки df2ed4841a9453ca
// Назначение: тест VoteTruth_Fb2oo2DAAI_MatchesTable набора FB_VoteTruth_Test.
// Автор:      kr0nsch; код — генератор cemgen
// Версия:     1.0.0
// Документ:   docs/DESIGN.md, раздел «10. Генератор cemgen»; docs/cause_effect_matrix.md
// ВНИМАНИЕ:   код демонстрационный и не предназначен для систем безопасности. Реальная ПАЗ требует
//             определения SIL, сертифицированных аппаратных и программных средств и валидации по
//             ГОСТ Р МЭК 61511.
// FB_Voting, схема 2oo2, политика DegradeAvailable, аналоговые каналы: все 64 сочетаний «требование ×
// достоверность × запрос байпаса» совпадают с таблицей TT_FB_2OO2_DA_AI. На строку — два вызова одного
// экземпляра: без запросов байпаса (сброс байпасов прошлой строки) и с полной строкой.
METHOD PRIVATE Fb2oo2DAAIMatchesTable
VAR
    fbTime     : PL.FB_FakeTime;   // время не меняется
    fbVote     : FB_Voting;        // ФБ под тестом, один экземпляр на все строки
    stCfg      : ST_VotingCfg;     // конфигурация теста уровня 2
    stIn       : ST_VoteIn;        // входы строки
    stCmd      : ST_VoteCmd;       // запросы байпаса строки
    uiRow      : UINT;             // строка таблицы
    bAct       : BYTE;             // фактический байт результата
    bExp       : BYTE;             // ожидаемый байт из таблицы
    xMiss      : BOOL;             // строка не совпала
    xFirst     : BOOL;             // первая несовпавшая строка
    uiMismatch : UINT;             // несовпавших строк
    uiFirstRow : UINT;             // первая несовпавшая строка
    bFirstExp  : BYTE;             // ожидаемый байт первой несовпавшей строки
    bFirstAct  : BYTE;             // фактический байт первой несовпавшей строки
END_VAR

(* ---- Fb2oo2DAAIMatchesTable.method.impl.st ---- *)
// AUTO-GENERATED by cemgen 1.0.0 — не редактировать: правьте матрицу и запустите
//   python -m cemgen generate <файл матрицы .csv или .xlsx>
// Матрица: SIS-V101-CEM, объект V-101, ревизия B от 2026-10-19, SHA-256 сетки df2ed4841a9453ca
coUnit.TEST('VoteTruth_Fb2oo2DAAI_MatchesTable');
stCfg.eArch := E_VoteArch.Vote2oo2;
stCfg.ePolicy := E_DegradePolicy.DegradeAvailable;
stCfg.eInput := E_SisInputKind.Analog;
stCfg.xDiHealthy := TRUE;
stCfg.eLimitDir := E_LimitDir.High;
stCfg.rTripLimit_eu := 50.0;
stCfg.rHyst_eu := 0.0;
stCfg.rDiscrepancyMax_eu := 0.0;
stCfg.tDiscrepancyDelay := T#0S;
stCfg.tBypassMax := T#1H;
stCfg.uiMaxBypass := 1;
FOR uiRow := 0 TO 63 DO
    RowInputs(uiRow := uiRow, uiChannels := 2, xBypass := FALSE, stIn := stIn, stCmd := stCmd);
    fbVote(stIn := stIn, stCmd := stCmd, stCfg := stCfg, xBypassPermit := TRUE, uiCause := 1,
        itfTime := fbTime);
    RowInputs(uiRow := uiRow, uiChannels := 2, xBypass := TRUE, stIn := stIn, stCmd := stCmd);
    fbVote(stIn := stIn, stCmd := stCmd, stCfg := stCfg, xBypassPermit := TRUE, uiCause := 1,
        itfTime := fbTime);
    bAct := EncodeFb(xTrip := fbVote.xTrip, stSts := fbVote.stSts);
    bExp := GVL_VoteTruthTable.TT_FB_2OO2_DA_AI[uiRow];
    xMiss := bAct <> bExp;
    xFirst := xMiss AND uiMismatch = 0;
    uiFirstRow := SEL(xFirst, uiFirstRow, uiRow);
    bFirstExp := SEL(xFirst, bFirstExp, bExp);
    bFirstAct := SEL(xFirst, bFirstAct, bAct);
    uiMismatch := uiMismatch + BOOL_TO_UINT(xMiss);
END_FOR
AssertEquals_UINT(Expected := 0, Actual := uiMismatch,
    Message := MismatchText(sTable := 'TT_FB_2OO2_DA_AI', uiRow := uiFirstRow, bExpected := bFirstExp,
        bActual := bFirstAct));
coUnit.TEST_FINISHED();

(* ---- Fb2oo2DADIMatchesTable.method.decl.st ---- *)
// AUTO-GENERATED by cemgen 1.0.0 — не редактировать: правьте матрицу и запустите
//   python -m cemgen generate <файл матрицы .csv или .xlsx>
// Матрица: SIS-V101-CEM, объект V-101, ревизия B от 2026-10-19, SHA-256 сетки df2ed4841a9453ca
// Назначение: тест VoteTruth_Fb2oo2DADI_MatchesTable набора FB_VoteTruth_Test.
// Автор:      kr0nsch; код — генератор cemgen
// Версия:     1.0.0
// Документ:   docs/DESIGN.md, раздел «10. Генератор cemgen»; docs/cause_effect_matrix.md
// ВНИМАНИЕ:   код демонстрационный и не предназначен для систем безопасности. Реальная ПАЗ требует
//             определения SIL, сертифицированных аппаратных и программных средств и валидации по
//             ГОСТ Р МЭК 61511.
// FB_Voting, схема 2oo2, политика DegradeAvailable, дискретные каналы: все 64 сочетаний «требование ×
// достоверность × запрос байпаса» совпадают с таблицей TT_FB_2OO2_DA_DI. На строку — два вызова одного
// экземпляра: без запросов байпаса (сброс байпасов прошлой строки) и с полной строкой.
METHOD PRIVATE Fb2oo2DADIMatchesTable
VAR
    fbTime     : PL.FB_FakeTime;   // время не меняется
    fbVote     : FB_Voting;        // ФБ под тестом, один экземпляр на все строки
    stCfg      : ST_VotingCfg;     // конфигурация теста уровня 2
    stIn       : ST_VoteIn;        // входы строки
    stCmd      : ST_VoteCmd;       // запросы байпаса строки
    uiRow      : UINT;             // строка таблицы
    bAct       : BYTE;             // фактический байт результата
    bExp       : BYTE;             // ожидаемый байт из таблицы
    xMiss      : BOOL;             // строка не совпала
    xFirst     : BOOL;             // первая несовпавшая строка
    uiMismatch : UINT;             // несовпавших строк
    uiFirstRow : UINT;             // первая несовпавшая строка
    bFirstExp  : BYTE;             // ожидаемый байт первой несовпавшей строки
    bFirstAct  : BYTE;             // фактический байт первой несовпавшей строки
END_VAR
